(* Logix 5000 project; controller TFF vendor 1 type 14 code 107 rev 34.11; software revision 34.03; part 21 of 36 *)
(* tags used below, declared in another part *)
   Address : DINT;   // Temp Address
   Config : Configuration;   // Index Array used in configuration routines
   AI101 : ALIAS FOR AnalogPoint[10];   // Filtrate Conductivity
   AlarmAnalog : AlarmAnalog[50];   // Analog Alarm Array
   AnalogOutput : AnalogOutput[25];   // Analog Output Array
   AnalogPoint : AnalogInput[50];   // Analog Input Array
   Concentration : Concentration;
   ControlLoop : ControlLoop[20];   // Control Loop Array
   ControlLoop_FeedBagLevel : ALIAS FOR ControlLoop[2];   // Feed Bag Level Control Loop
   ControlLoop_FeedPump : ALIAS FOR ControlLoop[1];   // Feed Pump Control Loop
   Diafiltration : Diafiltration;
   DigitalPoint : DigitalPoint[150];   // Digital Point Array
   Drive : Drive[11];   // Drives Array
   FI003 : ALIAS FOR AnalogPoint[17];
   FlowPath : FlowPath[64];   // Flow Path Array
   FlowPathControl : FlowPathControl;   // Flow Path Control
   FQ_Conc : ALIAS FOR Totalizer[0];   // Concentration Totalizer
   FQ_Diaf : ALIAS FOR Totalizer[1];   // DiafiltrationTotalizer
   Mixer : Mixer;   // Mixer config. structure
   Options : Options;   // Options List
   PCV001 : ALIAS FOR AnalogPoint[3];   // Retentate Pressure Control Valve Position
   PCV101 : ALIAS FOR AnalogPoint[4];   // Filtrate Pressure Control Valve Position
   Phase : Phases[6];   // Phase Control Array
   Phase0_Totalizer_Feed : ALIAS FOR PhaseTotalizer[0];   // Phase 0 Total Feed
   Phase0_Totalizer_Filtrate : ALIAS FOR PhaseTotalizer[6];   // Phase 0 Total Filtrate
   Phase0_Totalizer_Retentate : ALIAS FOR PhaseTotalizer[12];   // Phase 0 Total Retentate
   Phase1_Totalizer_Feed : ALIAS FOR PhaseTotalizer[1];   // Phase 1 Total Feed
   Phase1_Totalizer_Filtrate : ALIAS FOR PhaseTotalizer[7];   // Phase 1 Total Filtrate
   Phase1_Totalizer_Retentate : ALIAS FOR PhaseTotalizer[13];   // Phase 1 Total Retentate
   Phase2_Totalizer_Feed : ALIAS FOR PhaseTotalizer[2];   // Phase 2 Total Feed
   Phase2_Totalizer_Filtrate : ALIAS FOR PhaseTotalizer[8];   // Phase 2 Total Filtrate
   Phase2_Totalizer_Retentate : ALIAS FOR PhaseTotalizer[14];   // Phase 2 Total Retentate
   Phase3_Totalizer_Feed : ALIAS FOR PhaseTotalizer[3];   // Phase 3 Total Feed
   Phase3_Totalizer_Filtrate : ALIAS FOR PhaseTotalizer[9];   // Phase 3 Total Filtrate
   Phase3_Totalizer_Retentate : ALIAS FOR PhaseTotalizer[15];   // Phase 3 Total Retentate
   Phase4_Totalizer_Feed : ALIAS FOR PhaseTotalizer[4];   // Phase 4 Total Feed
   Phase4_Totalizer_Filtrate : ALIAS FOR PhaseTotalizer[10];   // Phase 4 Total Filtrate
   Phase4_Totalizer_Retentate : ALIAS FOR PhaseTotalizer[16];   // Phase 4 Total Retentate
   Phase5_Totalizer_Feed : ALIAS FOR PhaseTotalizer[5];   // Phase 5 Total Feed
   Phase5_Totalizer_Filtrate : ALIAS FOR PhaseTotalizer[11];   // Phase 5 Total Filtrate
   Phase5_Totalizer_Retentate : ALIAS FOR PhaseTotalizer[17];   // Phase 5 Total Retentate
   Rack_Murr_Node4_Instrum_TFF1 : IO_Station;   // Status of Node 4 Instrum TFF1
   Rack_Murr_Node4_Instrum_TFF2 : IO_Station;   // Status of Node 4 Instrum TFF2
   Rack_Murr_Node4_Instrum_TFF3 : IO_Station;   // Status of Node 4 Instrum TFF3
   Rack_Murr_Node4_Instrum_TFF4 : IO_Station;   // Status of Node 4 Instrum TFF4
   Rack_Murr_Node4_Instrum_TFF5 : IO_Station;   // Status of Node 4 Instrum TFF5
   Rack_Murr_Node5_Tank100 : IO_Station;   // Status of Node 5 Tank 100L
   Rack_Murr_Node5_Tank250 : IO_Station;   // Status of Node 5 Tank 250L
   Rack_Murr_Node5_Tank50 : IO_Station;   // Status of Node 5 Tank 50L
   SIC001 : ALIAS FOR Drive[1];   // Feed Pump
   SIC002 : ALIAS FOR Drive[2];   // Transfer Pump
   SIC003 : ALIAS FOR Drive[3];   // Mixer
   SysControl : SysControl;   // General system status and command
   Tank : TankManagement;   // Tank Management
   ThisSystem : SystemType;
   Valve : Valve[100];   // Valve Array
   ValveControl : ValveControl;   // Valve Control
   XV001 : ALIAS FOR Valve[0];   // XV001
   XV002 : ALIAS FOR Valve[1];   // XV002
   XV003 : ALIAS FOR Valve[2];   // XV003
   XV004 : ALIAS FOR Valve[3];   // XV004
   XV005 : ALIAS FOR Valve[4];   // XV005
   XV006 : ALIAS FOR Valve[19];
   XV007 : ALIAS FOR Valve[20];
   XV102 : ALIAS FOR Valve[5];   // XV102
   XV401 : ALIAS FOR Valve[6];   // XV401
   XV402 : ALIAS FOR Valve[7];   // XV402
   XV403 : ALIAS FOR Valve[15];
   XV404 : ALIAS FOR Valve[16];
   XV405 : ALIAS FOR Valve[17];
   XV406 : ALIAS FOR Valve[18];
   XV411 : ALIAS FOR Valve[8];   // XV411
   XV421 : ALIAS FOR Valve[9];   // XV421
   XV431 : ALIAS FOR Valve[10];   // XV431
   XV441 : ALIAS FOR Valve[11];   // XV441
   XV501 : ALIAS FOR Valve[12];   // XV501
   XV502 : ALIAS FOR Valve[13];   // XV502
   XV901 : ALIAS FOR Valve[14];   // XV901
(* Process, continued *)

ROUTINE Config_Drive   (* structured text *)
   (* ==========================================================
   	Config Drive : Configure Drive Structure (for Pumps)
   
   	List of treatments
   		- Drive[1] : Feed Pump SIC001
   		- Drive[2] : Transfer Pump SIC002
   		- Drive[3] : Mixer SIC003
   		- Reset Loop : Set to 0 the Drive[0 and 4 to 10].EnableCfg
   
   -----------------------------------------------------------------------------------------------------------------------------------------------------
   	History
   		2019-AUG-13 - ACTEMIUM - B. Roch - Initial version for Candidate Release 3.00.00.00.a
   ============================================================*)
   
   
   (*Drive[1] : Feed Pump SIC001
   ============================================================*)
   Config.IndexDr := 1 ;
   Drive[1].EnableCfg := 1 ;
   Drive[1].OutputAddress := 3 ;
   Drive[1].InputAddress := 0 ;
   Drive[1].RunInput := 0 ;
   Drive[1].InterlockTimer.PRE := 1000 ;
   Drive[1].ReverseCfg := 0 ;
   Drive[1].DirectionAddress := 0 ;
   
   (*Drive[2] : Transfer Pump SIC002
   ============================================================*)
   Drive[2].EnableCfg := 1 ;
   Drive[2].OutputAddress := 4 ;
   Drive[2].InputAddress := 0 ;
   Drive[2].RunInput := 0 ;
   Drive[2].InterlockTimer.PRE := 1000 ;
   Drive[2].ReverseCfg := 0 ;
   Drive[2].DirectionAddress := 0 ;
   
   (*Drive[3] : Mixer SIC003
   ============================================================*)
   Drive[3].EnableCfg := 1 ;
   Drive[3].OutputAddress := 6 ;
   Drive[3].InputAddress := 0 ;
   Drive[3].RunInput := 0 ;
   Drive[3].InterlockTimer.PRE := 1000 ;
   Drive[3].ReverseCfg := 0 ;
   Drive[3].DirectionAddress := 0 ;
   
   (*Reset Loop : Set to 0 the Drive[0 and 4 to 10].EnableCfg
   ============================================================*)
   for Config.IndexDr := 0 to 10 by 1 do
   	if Config.IndexDr = 0 or Config.IndexDr >= 4 then
   		Drive[Config.IndexDr].EnableCfg := 0 ;
   	End_if ;
   End_for ;
END_ROUTINE

ROUTINE Config_Flowpath   (* structured text *)
   (* =======================================================================
   	Config Flowpath : Configure predifined flowpath
   
   	List of treatments
   		- Critical
   		- Inlets
   		- Flush
   		- Drain
   		- Process
   		- Product Recovery
   		- Open All Main Valve
   		- Close All Main Valve
   		- Open All Valve (reserved)
   		- Close All Valve (reserved)
   		- Reset Loop : Set to 0 the mask and truth of Flowpath[36 to 60]
   
   -----------------------------------------------------------------------------------------------------------------------------------------------------
   	History
   		2019-AUG-13 - ACTEMIUM - B. Roch - Initial version for Candidate Release 3.00.00.00.a
   		2019-SEP-09 - ACTEMIUM - Q. Spindler - Modifications for Candidate Release 3.00.00.00.c
   					- Remove Flush and Drain from the Open all valve and close all valves Flowpath
   		2020-SEP-30 - Merck - Q.Spindler - Modifications for Candidate Release 3.00.00.01.a
   					- Modify flowpath for Closed flowpath option
   					- Add Flexware installation flowpath
   		2023-MAR-03 - Merck - Q.Spindler - Modifications for Candidate Release 3.02.00.00.a
   					- Add Remove TF3S/Closed FP Valves from masks if not enabled
   =========================================================================*)
   
   (* Max flowpath number use as terminal value in loop
   =========================================================================*)
   FlowPathControl.MaxFlowPath := 63 ;
   
   (* Critical
   =========================================================================*)
   (* Critical *)
   
   	FlowPath[2].Mask1 := 2097151 ;
   	FlowPath[2].Mask2 := 0 ;
   	FlowPath[2].Mask3 := 0 ;
   	FlowPath[2].Mask4 := 0 ;
   	FlowPath[2].DrainMask := 1 ;
   	FlowPath[2].FlushMask := 1 ;
   	FlowPath[2].Truth1 := 524299 ;
   	FlowPath[2].Truth2 := 0 ;
   	FlowPath[2].Truth3 := 0 ;
   	FlowPath[2].Truth4 := 0 ;
   	FlowPath[2].DrainTruth := 0 ;
   	FlowPath[2].FlushTruth := 0 ;
   
   
   (* Inlets
   =========================================================================*)
   	(* All Source Valves Open *)
   	FlowPath[3].Mask1 := 1052608 ;
   	FlowPath[3].Mask2 := 0 ;
   	FlowPath[3].Mask3 := 0 ;
   	FlowPath[3].Mask4 := 0 ;
   	FlowPath[3].DrainMask := 0 ;
   	FlowPath[3].FlushMask := 0 ;
   	FlowPath[3].Truth1 := 1052608 ;
   	FlowPath[3].Truth2 := 0 ;
   	FlowPath[3].Truth3 := 0 ;
   	FlowPath[3].Truth4 := 0 ;
   	FlowPath[3].DrainTruth := 0 ;
   	FlowPath[3].FlushTruth := 0 ;
   
   	(* All Source Valves Closed *)
   	FlowPath[4].Mask1 := 1052608 ;
   	FlowPath[4].Mask2 := 0 ;
   	FlowPath[4].Mask3 := 0 ;
   	FlowPath[4].Mask4 := 0 ;
   	FlowPath[4].DrainMask := 0 ;
   	FlowPath[4].FlushMask := 0 ;
   	FlowPath[4].Truth1 := 0 ;
   	FlowPath[4].Truth2 := 0 ;
   	FlowPath[4].Truth3 := 0 ;
   	FlowPath[4].Truth4 := 0 ;
   	FlowPath[4].DrainTruth := 0 ;
   	FlowPath[4].FlushTruth := 0 ;
   
   	(* Feed Source Open *)
   	FlowPath[5].Mask1 := 2068416 ;
   	FlowPath[5].Mask2 := 0 ;
   	FlowPath[5].Mask3 := 0 ;
   	FlowPath[5].Mask4 := 0 ;
   	FlowPath[5].DrainMask := 0 ;
   	FlowPath[5].FlushMask := 0 ;
   	FlowPath[5].Truth1 := 256 ;
   	FlowPath[5].Truth2 := 0 ;
   	FlowPath[5].Truth3 := 0 ;
   	FlowPath[5].Truth4 := 0 ;
   	FlowPath[5].DrainTruth := 0 ;
   	FlowPath[5].FlushTruth := 0 ;
   
   	(* Buffer Source Open *)
   	FlowPath[6].Mask1 := 2068416 ;
   	FlowPath[6].Mask2 := 0 ;
   	FlowPath[6].Mask3 := 0 ;
   	FlowPath[6].Mask4 := 0 ;
   	FlowPath[6].DrainMask := 0 ;
   	FlowPath[6].FlushMask := 0 ;
   	FlowPath[6].Truth1 := 576 ;
   	FlowPath[6].Truth2 := 0 ;
   	FlowPath[6].Truth3 := 0 ;
   	FlowPath[6].Truth4 := 0 ;
   	FlowPath[6].DrainTruth := 0 ;
   	FlowPath[6].FlushTruth := 0 ;
   
   	(* Caustic Source Open *)
   	FlowPath[7].Mask1 := 2068416 ;
   	FlowPath[7].Mask2 := 0 ;
   	FlowPath[7].Mask3 := 0 ;
   	FlowPath[7].Mask4 := 0 ;
   	FlowPath[7].DrainMask := 0 ;
   	FlowPath[7].FlushMask := 0 ;
   	FlowPath[7].Truth1 := 1088 ;
   	FlowPath[7].Truth2 := 0 ;
   	FlowPath[7].Truth3 := 0 ;
   	FlowPath[7].Truth4 := 0 ;
   	FlowPath[7].DrainTruth := 0 ;
   	FlowPath[7].FlushTruth := 0 ;
   
   	(* Water Source Open *)
   	FlowPath[8].Mask1 := 2068416 ;
   	FlowPath[8].Mask2 := 0 ;
   	FlowPath[8].Mask3 := 0 ;
   	FlowPath[8].Mask4 := 0 ;
   	FlowPath[8].DrainMask := 0 ;
   	FlowPath[8].FlushMask := 0 ;
   	FlowPath[8].Truth1 := 2112 ;
   	FlowPath[8].Truth2 := 0 ;
   	FlowPath[8].Truth3 := 0 ;
   	FlowPath[8].Truth4 := 0 ;
   	FlowPath[8].DrainTruth := 0 ;
   	FlowPath[8].FlushTruth := 0 ;
   
   	(* Air Source Open *)
   	FlowPath[9].Mask1 := 2068416 ;
   	FlowPath[9].Mask2 := 0 ;
   	FlowPath[9].Mask3 := 0 ;
   	FlowPath[9].Mask4 := 0 ;
   	FlowPath[9].DrainMask := 0 ;
   	FlowPath[9].FlushMask := 0 ;
   	FlowPath[9].Truth1 := 192 ;
   	FlowPath[9].Truth2 := 0 ;
   	FlowPath[9].Truth3 := 0 ;
   	FlowPath[9].Truth4 := 0 ;
   	FlowPath[9].DrainTruth := 0 ;
   	FlowPath[9].FlushTruth := 0 ;
   
   
   	(* Flush
   =========================================================================*)
   	(* Single Pass Flush (from inlet manifold) *)
   	FlowPath[10].Mask1 := 1044543 ;
   	FlowPath[10].Mask2 := 0 ;
   	FlowPath[10].Mask3 := 0 ;
   	FlowPath[10].Mask4 := 0 ;
   	FlowPath[10].DrainMask := 1 ;
   	FlowPath[10].FlushMask := 1 ;
   	FlowPath[10].Truth1 := 393227 ;
   	FlowPath[10].Truth2 := 0 ;
   	FlowPath[10].Truth3 := 0 ;
   	FlowPath[10].Truth4 := 0 ;
   	FlowPath[10].DrainTruth := 1 ;
   	FlowPath[10].FlushTruth := 1 ;
   
   	(* Single Pass Flush (from recycle bag) *)
   	FlowPath[11].Mask1 := 1044543 ;
   	FlowPath[11].Mask2 := 0 ;
   	FlowPath[11].Mask3 := 0 ;
   	FlowPath[11].Mask4 := 0 ;
   	FlowPath[11].DrainMask := 1 ;
   	FlowPath[11].FlushMask := 1 ;
   	FlowPath[11].Truth1 := 65547 ;
   	FlowPath[11].Truth2 := 0 ;
   	FlowPath[11].Truth3 := 0 ;
   	FlowPath[11].Truth4 := 0 ;
   	FlowPath[11].DrainTruth := 1 ;
   	FlowPath[11].FlushTruth := 0 ;
   
   
   	(* Drain
   =========================================================================*)
   	(* System Drain (without recycle bag) *)
   	FlowPath[12].Mask1 := 1044543 ;
   	FlowPath[12].Mask2 := 0 ;
   	FlowPath[12].Mask3 := 0 ;
   	FlowPath[12].Mask4 := 0 ;
   	FlowPath[12].DrainMask := 1 ;
   	FlowPath[12].FlushMask := 1 ;
   	FlowPath[12].Truth1 := 409647 ;
   	FlowPath[12].Truth2 := 0 ;
   	FlowPath[12].Truth3 := 0 ;
   	FlowPath[12].Truth4 := 0 ;
   	FlowPath[12].DrainTruth := 1 ;
   	FlowPath[12].FlushTruth := 1 ;
   
   	(* System Drain (from recycle bag) *)
   	FlowPath[13].Mask1 := 1044543 ;
   	FlowPath[13].Mask2 := 0 ;
   	FlowPath[13].Mask3 := 0 ;
   	FlowPath[13].Mask4 := 0 ;
   	FlowPath[13].DrainMask := 1 ;
   	FlowPath[13].FlushMask := 1 ;
   	FlowPath[13].Truth1 := 81983 ;
   	FlowPath[13].Truth2 := 0 ;
   	FlowPath[13].Truth3 := 0 ;
   	FlowPath[13].Truth4 := 0 ;
   	FlowPath[13].DrainTruth := 1 ;
   	FlowPath[13].FlushTruth := 0 ;
   
   
   	(* Process
   =========================================================================*)
   	(* Membrane Soak *)
   	FlowPath[14].Mask1 := 1044543 ;
   	FlowPath[14].Mask2 := 0 ;
   	FlowPath[14].Mask3 := 0 ;
   	FlowPath[14].Mask4 := 0 ;
   	FlowPath[14].DrainMask := 1 ;
   	FlowPath[14].FlushMask := 1 ;
   	FlowPath[14].Truth1 := 65539 ;
   	FlowPath[14].Truth2 := 0 ;
   	FlowPath[14].Truth3 := 0 ;
   	FlowPath[14].Truth4 := 0 ;
   	FlowPath[14].DrainTruth := 0 ;
   	FlowPath[14].FlushTruth := 0 ;
   
   	(* Integrity Test *)
   	FlowPath[15].Mask1 := 1044543 ;
   	FlowPath[15].Mask2 := 0 ;
   	FlowPath[15].Mask3 := 0 ;
   	FlowPath[15].Mask4 := 0 ;
   	FlowPath[15].DrainMask := 1 ;
   	FlowPath[15].FlushMask := 1 ;
   	FlowPath[15].Truth1 := 48 ;
   	FlowPath[15].Truth2 := 0 ;
   	FlowPath[15].Truth3 := 0 ;
   	FlowPath[15].Truth4 := 0 ;
   	FlowPath[15].DrainTruth := 0 ;
   	FlowPath[15].FlushTruth := 0 ;
   
   	(* Recycle Bag Fill *)
   	FlowPath[16].Mask1 := 1044543 ;
   	FlowPath[16].Mask2 := 0 ;
   	FlowPath[16].Mask3 := 0 ;
   	FlowPath[16].Mask4 := 0 ;
   	FlowPath[16].DrainMask := 1 ;
   	FlowPath[16].FlushMask := 1 ;
   	FlowPath[16].Truth1 := 524312 ;
   	FlowPath[16].Truth2 := 0 ;
   	FlowPath[16].Truth3 := 0 ;
   	FlowPath[16].Truth4 := 0 ;
   	FlowPath[16].DrainTruth := 0 ;
   	FlowPath[16].FlushTruth := 0 ;
   
   	(* Recycle Bag Drain *)
   	FlowPath[17].Mask1 := 1044543 ;
   	FlowPath[17].Mask2 := 0 ;
   	FlowPath[17].Mask3 := 0 ;
   	FlowPath[17].Mask4 := 0 ;
   	FlowPath[17].DrainMask := 1 ;
   	FlowPath[17].FlushMask := 1 ;
   	FlowPath[17].Truth1 := 81925 ;
   	FlowPath[17].Truth2 := 0 ;
   	FlowPath[17].Truth3 := 0 ;
   	FlowPath[17].Truth4 := 0 ;
   	FlowPath[17].DrainTruth := 0 ;
   	FlowPath[17].FlushTruth := 0 ;
   
   	(* Recovery Filter Flush *)
   	FlowPath[18].Mask1 := 1044543 ;
   	FlowPath[18].Mask2 := 0 ;
   	FlowPath[18].Mask3 := 0 ;
   	FlowPath[18].Mask4 := 0 ;
   	FlowPath[18].DrainMask := 1 ;
   	FlowPath[18].FlushMask := 1 ;
   	FlowPath[18].Truth1 := 65541 ;
   	FlowPath[18].Truth2 := 0 ;
   	FlowPath[18].Truth3 := 0 ;
   	FlowPath[18].Truth4 := 0 ;
   	FlowPath[18].DrainTruth := 0 ;
   	FlowPath[18].FlushTruth := 0 ;
   
   	(* Batch UF or Membrane Recycle *)
   	FlowPath[19].Mask1 := 1044543 ;
   	FlowPath[19].Mask2 := 0 ;
   	FlowPath[19].Mask3 := 0 ;
   	FlowPath[19].Mask4 := 0 ;
   	FlowPath[19].DrainMask := 1 ;
   	FlowPath[19].FlushMask := 1 ;
   	FlowPath[19].Truth1 := 589835 ;
   	FlowPath[19].Truth2 := 0 ;
   	FlowPath[19].Truth3 := 0 ;
   	FlowPath[19].Truth4 := 0 ;
   	FlowPath[19].DrainTruth := 0 ;
   	FlowPath[19].FlushTruth := 0 ;
   
   	(* Fed Batch UF or Diafiltration *)
   	FlowPath[20].Mask1 := 1044543 ;
   	FlowPath[20].Mask2 := 0 ;
   	FlowPath[20].Mask3 := 0 ;
   	FlowPath[20].Mask4 := 0 ;
   	FlowPath[20].DrainMask := 1 ;
   	FlowPath[20].FlushMask := 1 ;
   	FlowPath[20].Truth1 := 589851 ;
   	FlowPath[20].Truth2 := 0 ;
   	FlowPath[20].Truth3 := 0 ;
   	FlowPath[20].Truth4 := 0 ;
   	FlowPath[20].DrainTruth := 0 ;
   	FlowPath[20].FlushTruth := 0 ;
   
   
   	(* Product Recovery
   =========================================================================*)
   	(* Product Recovery 1&3 - Empty Recycle Bag (TF2S) *)
   	FlowPath[21].Mask1 := 1032255 ;
   	FlowPath[21].Mask2 := 0 ;
   	FlowPath[21].Mask3 := 0 ;
   	FlowPath[21].Mask4 := 0 ;
   	FlowPath[21].DrainMask := 1 ;
   	FlowPath[21].FlushMask := 1 ;
   	FlowPath[21].Truth1 := 65541 ;
   	FlowPath[21].Truth2 := 0 ;
   	FlowPath[21].Truth3 := 0 ;
   	FlowPath[21].Truth4 := 0 ;
   	FlowPath[21].DrainTruth := 0 ;
   	FlowPath[21].FlushTruth := 0 ;
   
   	(* Product Recovery 2 - Empty Retentate Line (TF2S) *)
   	FlowPath[22].Mask1 := 1032255 ;
   	FlowPath[22].Mask2 := 0 ;
   	FlowPath[22].Mask3 := 0 ;
   	FlowPath[22].Mask4 := 0 ;
   	FlowPath[22].DrainMask := 1 ;
   	FlowPath[22].FlushMask := 1 ;
   	FlowPath[22].Truth1 := 524312 ;
   	FlowPath[22].Truth2 := 0 ;
   	FlowPath[22].Truth3 := 0 ;
   	FlowPath[22].Truth4 := 0 ;
   	FlowPath[22].DrainTruth := 0 ;
   	FlowPath[22].FlushTruth := 0 ;
   
   	(* Product Recovery 4 - Empty Membranes (TF2S) *)
   	FlowPath[23].Mask1 := 1032255 ;
   	FlowPath[23].Mask2 := 0 ;
   	FlowPath[23].Mask3 := 0 ;
   	FlowPath[23].Mask4 := 0 ;
   	FlowPath[23].DrainMask := 1 ;
   	FlowPath[23].FlushMask := 1 ;
   	FlowPath[23].Truth1 := 22 ;
   	FlowPath[23].Truth2 := 0 ;
   	FlowPath[23].Truth3 := 0 ;
   	FlowPath[23].Truth4 := 0 ;
   	FlowPath[23].DrainTruth := 0 ;
   	FlowPath[23].FlushTruth := 0 ;
   
   	(* Product Recovery 1&5 - Empty Recycle Bag (TF3S) *)
   	FlowPath[24].Mask1 := 1044543 ;
   	FlowPath[24].Mask2 := 0 ;
   	FlowPath[24].Mask3 := 0 ;
   	FlowPath[24].Mask4 := 0 ;
   	FlowPath[24].DrainMask := 1 ;
   	FlowPath[24].FlushMask := 1 ;
   	FlowPath[24].Truth1 := 65541 ;
   	FlowPath[24].Truth2 := 0 ;
   	FlowPath[24].Truth3 := 0 ;
   	FlowPath[24].Truth4 := 0 ;
   	FlowPath[24].DrainTruth := 0 ;
   	FlowPath[24].FlushTruth := 0 ;
   
   	(* Product Recovery 2 - Empty Membranes (TF3S) *)
   	FlowPath[25].Mask1 := 1044543 ;
   	FlowPath[25].Mask2 := 0 ;
   	FlowPath[25].Mask3 := 0 ;
   	FlowPath[25].Mask4 := 0 ;
   	FlowPath[25].DrainMask := 1 ;
   	FlowPath[25].FlushMask := 1 ;
   	FlowPath[25].Truth1 := 22 ;
   	FlowPath[25].Truth2 := 0 ;
   	FlowPath[25].Truth3 := 0 ;
   	FlowPath[25].Truth4 := 0 ;
   	FlowPath[25].DrainTruth := 0 ;
   	FlowPath[25].FlushTruth := 0 ;
   
   	(* Product Recovery 3&6 - Empty Bypass (TF3S) *)
   	FlowPath[26].Mask1 := 1044543 ;
   	FlowPath[26].Mask2 := 0 ;
   	FlowPath[26].Mask3 := 0 ;
   	FlowPath[26].Mask4 := 0 ;
   	FlowPath[26].DrainMask := 1 ;
   	FlowPath[26].FlushMask := 1 ;
   	FlowPath[26].Truth1 := 12310 ;
   	FlowPath[26].Truth2 := 0 ;
   	FlowPath[26].Truth3 := 0 ;
   	FlowPath[26].Truth4 := 0 ;
   	FlowPath[26].DrainTruth := 0 ;
   	FlowPath[26].FlushTruth := 0 ;
   
   	(* Product Recovery 4 - Empty Retentate Line (TF3S) *)
   	FlowPath[27].Mask1 := 1044543 ;
   	FlowPath[27].Mask2 := 0 ;
   	FlowPath[27].Mask3 := 0 ;
   	FlowPath[27].Mask4 := 0 ;
   	FlowPath[27].DrainMask := 1 ;
   	FlowPath[27].FlushMask := 1 ;
   	FlowPath[27].Truth1 := 524312 ;
   	FlowPath[27].Truth2 := 0 ;
   	FlowPath[27].Truth3 := 0 ;
   	FlowPath[27].Truth4 := 0 ;
   	FlowPath[27].DrainTruth := 0 ;
   	FlowPath[27].FlushTruth := 0 ;
   
   
   (* Open All Main Valve
   =========================================================================*)
   	(* All Main Flowpath Valves Open *)
   	FlowPath[28].Mask1 := 1044543 ;
   	FlowPath[28].Mask2 := 0 ;
   	FlowPath[28].Mask3 := 0 ;
   	FlowPath[28].Mask4 := 0 ;
   	FlowPath[28].DrainMask := 1 ;
   	FlowPath[28].FlushMask := 1 ;
   	FlowPath[28].Truth1 := 606271 ;
   	FlowPath[28].Truth2 := 0 ;
   	FlowPath[28].Truth3 := 0 ;
   	FlowPath[28].Truth4 := 0 ;
   	FlowPath[28].DrainTruth := 0 ;
   	FlowPath[28].FlushTruth := 0 ;
   
   
   (* Close All Main Valve
   =========================================================================*)
   	(* All Main Flowpath Valves Closed *)
   	FlowPath[29].Mask1 := 1044543 ;
   	FlowPath[29].Mask2 := 0 ;
   	FlowPath[29].Mask3 := 0 ;
   	FlowPath[29].Mask4 := 0 ;
   	FlowPath[29].DrainMask := 1 ;
   	FlowPath[29].FlushMask := 1 ;
   	FlowPath[29].Truth1 := 0 ;
   	FlowPath[29].Truth2 := 0 ;
   	FlowPath[29].Truth3 := 0 ;
   	FlowPath[29].Truth4 := 0 ;
   	FlowPath[29].DrainTruth := 0 ;
   	FlowPath[29].FlushTruth := 0 ;
   
   
   (* Flowpath from 30 to 34 are reserved for User *)
   
   	(* FlexWare Installation *)
   	FlowPath[35].Mask1 := 2068416 ;
   	FlowPath[35].Mask2 := 0 ;
   	FlowPath[35].Mask3 := 0 ;
   	FlowPath[35].Mask4 := 0 ;
   	FlowPath[35].DrainMask := 0 ;
   	FlowPath[35].FlushMask := 0 ;
   	FlowPath[35].Truth1 := 2068416 ;
   	FlowPath[35].Truth2 := 0 ;
   	FlowPath[35].Truth3 := 0 ;
   	FlowPath[35].Truth4 := 0 ;
   	FlowPath[35].DrainTruth := 0 ;
   	FlowPath[35].FlushTruth := 0 ;
   
   
   // Remove TF3S Valves from mask if not enabled
   IF NOT Options.TF3S THEN
   	FOR Config.IndexFlowpath := 2 to 29 by 1 do
   		FlowPath[Config.IndexFlowpath].Mask1.12 := 0 ; //XV501
   		FlowPath[Config.IndexFlowpath].Mask1.13 := 0 ; //XV502
   	End_for ;
   		FlowPath[35].Mask1.12 := 0 ; //XV501
   		FlowPath[35].Mask1.13 := 0 ; //XV502
   END_IF;
   
   // Remove Closed FP Valves from mask if not enabled
   IF NOT Options.ClosedFP THEN
   	FOR Config.IndexFlowpath := 2 to 29 by 1 do
   		FlowPath[Config.IndexFlowpath].Mask1.15 := 0 ; //XV403
   		FlowPath[Config.IndexFlowpath].Mask1.16 := 0 ; //XV404
   		FlowPath[Config.IndexFlowpath].Mask1.17 := 0 ; //XV405
   		FlowPath[Config.IndexFlowpath].Mask1.18 := 0 ; //XV406
   		FlowPath[Config.IndexFlowpath].Mask1.19 := 0 ; //XV006
   		FlowPath[Config.IndexFlowpath].Mask1.20 := 0 ; //XV007
   	End_for ;
   		FlowPath[35].Mask1.15 := 0 ; //XV403
   		FlowPath[35].Mask1.16 := 0 ; //XV404
   		FlowPath[35].Mask1.17 := 0 ; //XV405
   		FlowPath[35].Mask1.18 := 0 ; //XV406
   		FlowPath[35].Mask1.19 := 0 ; //XV006
   		FlowPath[35].Mask1.20 := 0 ; //XV007
   END_IF;
   
   
   (* Open All Valve (reserved)
   =========================================================================*)
   (* Open All Valve *)
   FlowPath[61].Mask1 := -1 ;
   FlowPath[61].Mask2 := 0 ;
   FlowPath[61].Mask3 := 0 ;
   FlowPath[61].Mask4 := 0 ;
   FlowPath[61].DrainMask := 0 ;
   FlowPath[61].FlushMask := 0 ;
   FlowPath[61].Truth1 := -1 ;
   FlowPath[61].Truth2 := 0 ;
   FlowPath[61].Truth3 := 0 ;
   FlowPath[61].Truth4 := 0 ;
   FlowPath[61].DrainTruth := 0 ;
   FlowPath[61].FlushTruth := 0 ;
   
   (* Close All Valve (reserved)
   =========================================================================*)
   (* Close All Valve *)
   FlowPath[62].Mask1 := -1 ;
   FlowPath[62].Mask2 := 0 ;
   FlowPath[62].Mask3 := 0 ;
   FlowPath[62].Mask4 := 0 ;
   FlowPath[62].DrainMask := 0 ;
   FlowPath[62].FlushMask := 0 ;
   FlowPath[62].Truth1 := 0 ;
   FlowPath[62].Truth2 := 0 ;
   FlowPath[62].Truth3 := 0 ;
   FlowPath[62].Truth4 := 0 ;
   FlowPath[62].DrainTruth := 0 ;
   FlowPath[62].FlushTruth := 0 ;
   
   (*Reset Loop : Set to 0 the Flowpath[36 to 60]
   ============================================================*)
   FOR Config.IndexFlowpath := 36 to 60 by 1 do
   	FlowPath[Config.IndexFlowpath].Mask1 := 0 ;
   	FlowPath[Config.IndexFlowpath].Mask2 := 0 ;
   	FlowPath[Config.IndexFlowpath].Mask3 := 0 ;
   	FlowPath[Config.IndexFlowpath].Mask4 := 0 ;
   	FlowPath[Config.IndexFlowpath].DrainMask := 0 ;
   	FlowPath[Config.IndexFlowpath].FlushMask := 0 ;
   	FlowPath[Config.IndexFlowpath].Truth1 := 0 ;
   	FlowPath[Config.IndexFlowpath].Truth2 := 0 ;
   	FlowPath[Config.IndexFlowpath].Truth3 := 0 ;
   	FlowPath[Config.IndexFlowpath].Truth4 := 0 ;
   	FlowPath[Config.IndexFlowpath].Status := 0 ;
   	FlowPath[Config.IndexFlowpath].DrainTruth := 0 ;
   	FlowPath[Config.IndexFlowpath].FlushTruth := 0 ;
   End_for ;
END_ROUTINE

ROUTINE Config_Options   (* structured text *)
   (* ==========================================================
   	Config Options : Configure Options
   
   	List of treatments
   		- Configure Instrum TFF options
   		- Configure Tank options
   		- Configure Flag for current installed clamshell
   
   -----------------------------------------------------------------------------------------------------------------------------------------------------
   	History
   		2019-AUG-13 - ACTEMIUM - B. Roch - Initial version for Candidate Release 3.00.00.00.a
   ============================================================*)
   
   (*Configure options if option Simulation mode is disabled*)
   If Not SysControl.Simulate_Options Then
   
   	(* Configure Instrum TFF options
   	Set options depending on which INSTRUM_TFF I/O device is active
   	============================================================*)
   
   	(*No Device Connected*)
   	IF NOT Rack_Murr_Node4_Instrum_TFF1.Node_Comm_Status AND NOT Rack_Murr_Node4_Instrum_TFF2.Node_Comm_Status AND NOT Rack_Murr_Node4_Instrum_TFF3.Node_Comm_Status AND NOT Rack_Murr_Node4_Instrum_TFF4.Node_Comm_Status AND NOT Rack_Murr_Node4_Instrum_TFF5.Node_Comm_Status THEN
   	Options.No_Device_Connected := 1 ;
   	Options.AI102_AI103 := 0 ;
   	Options.AI101 := 0 ;
   	Options.AI101_AI102_AI103 := 0 ;
   	Options.AI101_AI104 := 0 ;
   	Options.AI101_AI102_AI103_AI104 := 0 ;
   	END_IF;
   
   	(*UV Probe Device*)
   	IF Rack_Murr_Node4_Instrum_TFF1.Node_Comm_Status THEN
   	Options.No_Device_Connected := 0 ;
   	Options.AI102_AI103 := 1 ;
   	Options.AI101 := 0 ;
   	Options.AI101_AI102_AI103 := 0 ;
   	Options.AI101_AI104 := 0 ;
   	Options.AI101_AI102_AI103_AI104 := 0 ;
   	END_IF;
   
   	(*Conductivity*)
   	IF Rack_Murr_Node4_Instrum_TFF2.Node_Comm_Status THEN
   	Options.No_Device_Connected := 0 ;
   	Options.AI102_AI103 := 0 ;
   	Options.AI101 := 1 ;
   	Options.AI101_AI102_AI103 := 0 ;
   	Options.AI101_AI104 := 0 ;
   	Options.AI101_AI102_AI103_AI104 := 0 ;
   	END_IF;
   
   	(*UV and Conductivity*)
   	IF Rack_Murr_Node4_Instrum_TFF3.Node_Comm_Status THEN
   	Options.No_Device_Connected := 0 ;
   	Options.AI102_AI103 := 0 ;
   	Options.AI101 := 0 ;
   	Options.AI101_AI102_AI103 := 1 ;
   	Options.AI101_AI104 := 0 ;
   	Options.AI101_AI102_AI103_AI104 := 0 ;
   	END_IF;
   
   	(*Conductivity and pH*)
   	IF Rack_Murr_Node4_Instrum_TFF4.Node_Comm_Status THEN
   	Options.No_Device_Connected := 0 ;
   	Options.AI102_AI103 := 0 ;
   	Options.AI101 := 0 ;
   	Options.AI101_AI102_AI103 := 0 ;
   	Options.AI101_AI104 := 1 ;
   	Options.AI101_AI102_AI103_AI104 := 0 ;
   	END_IF;
   
   	(*UV and Conductivity and pH*)
   	IF Rack_Murr_Node4_Instrum_TFF5.Node_Comm_Status THEN
   	Options.No_Device_Connected := 0 ;
   	Options.AI102_AI103 := 0 ;
   	Options.AI101 := 0 ;
   	Options.AI101_AI102_AI103 := 0 ;
   	Options.AI101_AI104 := 0 ;
   	Options.AI101_AI102_AI103_AI104 := 1 ;
   	END_IF;
   
   	(* Configure Tank options
   	Set options depending on which TANK I/O device is active
   	============================================================*)
   
   	(*No Tank Connected*)
   	IF NOT Rack_Murr_Node5_Tank50.Node_Comm_Status AND NOT Rack_Murr_Node5_Tank100.Node_Comm_Status AND NOT Rack_Murr_Node5_Tank250.Node_Comm_Status THEN
   	Options.No_Tank := 1 ;
   	Options.Tank50 := 0 ;
   	Options.Tank100 := 0 ;
   	Options.Tank250 := 0 ;
   	Tank.Config.Option_Current := 0 ;
   	END_IF;
   
   	(*Tank 50*)
   	IF Rack_Murr_Node5_Tank50.Node_Comm_Status THEN
   	Options.No_Tank := 0 ;
   	Options.Tank50 := 1 ;
   	Options.Tank100 := 0 ;
   	Options.Tank250 := 0 ;
   	Tank.Config.Option_Current := 1 ;
   	END_IF;
   
   	(*Tank 100*)
   	IF Rack_Murr_Node5_Tank100.Node_Comm_Status THEN
   	Options.No_Tank := 0 ;
   	Options.Tank50 := 0 ;
   	Options.Tank100 := 1 ;
   	Options.Tank250 := 0 ;
   	Tank.Config.Option_Current := 2 ;
   	END_IF;
   
   	(*Tank 250*)
   	IF Rack_Murr_Node5_Tank250.Node_Comm_Status THEN
   	Options.No_Tank := 0 ;
   	Options.Tank50 := 0 ;
   	Options.Tank100 := 0 ;
   	Options.Tank250 := 1 ;
   	Tank.Config.Option_Current := 3 ;
   	END_IF;
   
   End_If;
   
   
   (*Simulate Tank Range*)
   IF Tank.Config.Simulate THEN
   
   	CASE	Tank.Config.Option_Simulate OF
   		0:	Options.No_Tank := 1 ;
   			Options.Tank50 := 0 ;
   			Options.Tank100 := 0 ;
   			Options.Tank250 := 0 ;
   			Tank.Config.Option_Current := 0 ;
   		1:	Options.No_Tank := 0 ;
   			Options.Tank50 := 1 ;
   			Options.Tank100 := 0 ;
   			Options.Tank250 := 0 ;
   			Tank.Config.Option_Current := 1 ;
   		2:	Options.No_Tank := 0 ;
   			Options.Tank50 := 0 ;
   			Options.Tank100 := 1 ;
   			Options.Tank250 := 0 ;
   			Tank.Config.Option_Current := 2 ;
   		3:	Options.No_Tank := 0 ;
   			Options.Tank50 := 0 ;
   			Options.Tank100 := 0 ;
   			Options.Tank250 := 1 ;
   			Tank.Config.Option_Current := 3 ;
   	ELSE 	Options.No_Tank := 1 ;
   			Options.Tank50 := 0 ;
   			Options.Tank100 := 0 ;
   			Options.Tank250 := 0 ;
   			Tank.Config.Option_Current := 0 ;
   	END_CASE;
   
   END_IF;
   
   (* Configure Flag for current installed clamshell
   Used to create the CCP Configuration file based on current clamshell
   ============================================================*)
   IF ThisSystem.MoldType = 123 THEN
   
   	Options.TF2S := 1 ;
   	Options.TF3S := 0 ;
   
   ELSIF ThisSystem.MoldType = 124 THEN
   
   	Options.TF3S := 1 ;
   	Options.TF2S := 0 ;
   
   END_IF;
END_ROUTINE

ROUTINE Config_Reset   (* structured text *)
// Set to 0  all settings
   (* ==========================================================
   	Config Reset : 	When config.reset command is activated,AnalogPoint, AlarmAnalog, AnalogOutput, Drive, DigitalPoint and Valve structure
   					are initialized to 0.
   
   	List of treatments
   		- AnalogPoint Structure reset [0] to [49]
   		- AlarmAnalog Structure reset [0] to [49]
   		- AnalogOutput Structure reset [0] to [24]
   		- Drive Structure reset [0] to [10]
   		- DigitalPoint Structure reset [0] to [149]
   		- Valve Structure reset [0] to [99]
   
   -----------------------------------------------------------------------------------------------------------------------------------------------------
   	History
   		2019-AUG-13 - ACTEMIUM - B. Roch - Initial version for Candidate Release 3.00.00.00.a
   ============================================================*)
   
   
   (*Structure Reset [0] to [149]
   ============================================================*)
   IF Config.Reset THEN
   	FOR Config.IndexReset := 0 TO 149 BY 1 Do
   		IF Config.IndexReset <= 49 THEN
   		(*AnalogPoint Structure Reset [0] to [49]
   		====================================================*)
   			AnalogPoint[Config.IndexReset].OutofRange := 0 ;
   			AnalogPoint[Config.IndexReset].FilterType := 0 ;
   			AnalogPoint[Config.IndexReset].AveragingTotal := 0 ;
   			AnalogPoint[Config.IndexReset].Address := 0 ;
   			AnalogPoint[Config.IndexReset].RawMin := 0 ;
   			AnalogPoint[Config.IndexReset].RawMax := 0 ;
   			AnalogPoint[Config.IndexReset].RawValue := 0 ;
   			AnalogPoint[Config.IndexReset].RawLowLimit := 0 ;
   			AnalogPoint[Config.IndexReset].RawHighLimit := 0 ;
   			AnalogPoint[Config.IndexReset].FilterUser := 0 ;
   			AnalogPoint[Config.IndexReset].FilteredRaw := 0 ;
   			AnalogPoint[Config.IndexReset].FilterActual := 0 ;
   			AnalogPoint[Config.IndexReset].ScaledMin := 0 ;
   			AnalogPoint[Config.IndexReset].ScaledMax := 0 ;
   			AnalogPoint[Config.IndexReset].RangeMin := 0 ;
   			AnalogPoint[Config.IndexReset].RangeMax := 0 ;
   			AnalogPoint[Config.IndexReset].RangeMinSave := 0 ;
   			AnalogPoint[Config.IndexReset].RangeMaxSave := 0 ;
   			AnalogPoint[Config.IndexReset].RealCfg := 0 ;
   			AnalogPoint[Config.IndexReset].EnableCfg := 0 ;
   			AnalogPoint[Config.IndexReset].OverrideCfg := 0 ;
   
   		(*AlarmAnalog Structure Reset [0] to [49]
   		====================================================*)
   			AlarmAnalog[Config.IndexReset].Override := 0 ;
   			AlarmAnalog[Config.IndexReset].Disable := 0 ;
   			AlarmAnalog[Config.IndexReset].LOLODisable := 0 ;
   			AlarmAnalog[Config.IndexReset].LODisable := 0 ;
   			AlarmAnalog[Config.IndexReset].HIDisable := 0 ;
   			AlarmAnalog[Config.IndexReset].HIHIDisable := 0 ;
   			AlarmAnalog[Config.IndexReset].HIHIEnable := 0 ;
   			AlarmAnalog[Config.IndexReset].FeedPumpEnable := 0 ;
   			AlarmAnalog[Config.IndexReset].FeedPumpTag := 0 ;
   			AlarmAnalog[Config.IndexReset].TransferPumpEnable := 0 ;
   			AlarmAnalog[Config.IndexReset].TransferPumpTag := 0 ;
   			AlarmAnalog[Config.IndexReset].LOLO := 0 ;
   			AlarmAnalog[Config.IndexReset].LO := 0 ;
   			AlarmAnalog[Config.IndexReset].HI := 0 ;
   			AlarmAnalog[Config.IndexReset].HIHI := 0 ;
   			AlarmAnalog[Config.IndexReset].LOLOTimer.PRE := 0 ;
   			AlarmAnalog[Config.IndexReset].LOTimer.PRE := 0 ;
   			AlarmAnalog[Config.IndexReset].HITimer.PRE := 0 ;
   			AlarmAnalog[Config.IndexReset].HIHITimer.PRE := 0 ;
   			AlarmAnalog[Config.IndexReset].EnableCfg := 0 ;
   		End_IF;
   
   		(*AnalogOutput Structure Reset [0] to [24]
   		====================================================*)
   		IF Config.IndexReset <= 24 THEN
   			AnalogOutput[Config.IndexReset].RawValue := 0 ;
   			AnalogOutput[Config.IndexReset].RawMin := 0 ;
   			AnalogOutput[Config.IndexReset].RawMax := 0 ;
   			AnalogOutput[Config.IndexReset].ScaledMin := 0 ;
   			AnalogOutput[Config.IndexReset].ScaledMax := 0 ;
   			AnalogOutput[Config.IndexReset].EnableCfg := 0 ;
   		End_IF;
   
   		(*Drive Structure Reset [0] to [10]
   		====================================================*)
   		IF Config.IndexReset <= 10 THEN
   			Drive[Config.IndexReset].OutputAddress := 0 ;
   			Drive[Config.IndexReset].InputAddress := 0 ;
   			Drive[Config.IndexReset].RunInput := 0 ;
   			Drive[Config.IndexReset].InterlockTimer.PRE := 0 ;
   			Drive[Config.IndexReset].EnableCfg := 0 ;
   			Drive[Config.IndexReset].ReverseCfg := 0 ;
   			Drive[Config.IndexReset].Direction := 0 ;
   			Drive[Config.IndexReset].DirectionAddress := 0 ;
   		End_IF;
   
   		IF Config.IndexReset <= 99 THEN
   				(*Valves Structure Reset [0] to [99]
   		====================================================*)
   		Valve[Config.IndexReset].ZSOpenEnable := 0 ;
   		Valve[Config.IndexReset].ZSCloseEnable := 0 ;
   		Valve[Config.IndexReset].ZSOverride := 0 ;
   		Valve[Config.IndexReset].FailState := 0 ;
   		Valve[Config.IndexReset].Ports := 0 ;
   		Valve[Config.IndexReset].EnableCfg := 0 ;
   		Valve[Config.IndexReset].StatusWord := 0 ;
   		Valve[Config.IndexReset].ZSOpenAddress := 0 ;
   		Valve[Config.IndexReset].ZSCloseAddress := 0 ;
   		Valve[Config.IndexReset].OutputAddress := 0 ;
   		Valve[Config.IndexReset].AlarmTimer.PRE := 0 ;
   		Valve[Config.IndexReset].AutoCloseTimer.PRE := 0 ;
   		End_IF;
   
   		(*DigitalPoint Structure Reset [0] to [149]
   		====================================================*)
   		DigitalPoint[Config.IndexReset].Override := 0 ;
   		DigitalPoint[Config.IndexReset].DelayTimer.PRE := 0 ;
   		DigitalPoint[Config.IndexReset].Priority := 0 ;
   		DigitalPoint[Config.IndexReset].EnableCfg := 0 ;
   		DigitalPoint[Config.IndexReset].ActiveStateCFg := 0 ;
   		DigitalPoint[Config.IndexReset].RealInputCfg := 0 ;
   		DigitalPoint[Config.IndexReset].InputAddressCfg := 0 ;
   		DigitalPoint[Config.IndexReset].AlarmCfg := 0 ;
   		DigitalPoint[Config.IndexReset].AlarmStateCfg := 0 ;
   		DigitalPoint[Config.IndexReset].OverrideCfg := 0 ;
   		DigitalPoint[Config.IndexReset].PriorityCfg := 0 ;
   		DigitalPoint[Config.IndexReset].Cond1Cfg := 0 ;
   		DigitalPoint[Config.IndexReset].Cond2Cfg := 0 ;
   		DigitalPoint[Config.IndexReset].FlashingInputCfg := 0 ;
   
   	END_FOR;
   End_IF;
   (*Reset config.reset to execute routine one time*)
   Config.Reset := 0;
END_ROUTINE

ROUTINE Config_Totalizers   (* structured text *)
   (* ==========================================================
   	Config Totalizers : Configure Totalizers Structure
   
   	List of treatments
   		- Phase 0 Totalizers
   		- Phase 1 Totalizers
   		- Phase 2 Totalizers
   		- Phase 3 Totalizers
   		- Phase 4 Totalizers
   		- Phase 5 Totalizers
   		- Concentration and Diafiltration Totalizers
   
   -----------------------------------------------------------------------------------------------------------------------------------------------------
   	History
   		2019-AUG-13 - ACTEMIUM - B. Roch - Initial version for Candidate Release 3.00.00.00.a
   		2020-SEP-29 - Merck - Q. Spindler - Modifications for Candidate Release 3.00.00.01.a
   					- Add Retentate totalizers
   		2020-NOV-24 - Merck - Q. Spindler - Modifications for Candidate Release 3.00.00.01.b
   					- Change Retentate Flowmeter option
   ============================================================*)
   
   
   (*Phase 0 Totalizers
   ============================================================*)
   Phase0_Totalizer_Feed.EnableCfg := 1 ;
   Phase0_Totalizer_Feed.SourceAddressCfg := 42 ;
   Phase0_Totalizer_Feed.SourceTypeCfg := 0 ;
   Phase0_Totalizer_Feed.PVscale := 60 ;
   
   
   IF Options.No_Filtrate_Measurement THEN
   	Phase0_Totalizer_Filtrate.EnableCfg := 0 ;
   ELSE
   	Phase0_Totalizer_Filtrate.EnableCfg := 1 ;
   END_IF;
   
   Phase0_Totalizer_Filtrate.SourceAddressCfg := 2 ;
   Phase0_Totalizer_Filtrate.SourceTypeCfg := 0 ;
   Phase0_Totalizer_Filtrate.PVscale := 60 ;
   
   IF Options.FI003 THEN
   	Phase0_Totalizer_Retentate.EnableCfg := 1 ;
   ELSE
   	Phase0_Totalizer_Retentate.EnableCfg := 0 ;
   END_IF;
   
   Phase0_Totalizer_Retentate.SourceAddressCfg := 17 ;
   Phase0_Totalizer_Retentate.SourceTypeCfg := 0 ;
   Phase0_Totalizer_Retentate.PVscale := 60 ;
   
   (*Phase 1 Totalizers
   ============================================================*)
   Phase1_Totalizer_Feed.EnableCfg := 1 ;
   Phase1_Totalizer_Feed.SourceAddressCfg := 42 ;
   Phase1_Totalizer_Feed.SourceTypeCfg := 0 ;
   Phase1_Totalizer_Feed.PVscale := 60 ;
   
   IF Options.No_Filtrate_Measurement THEN
   	Phase1_Totalizer_Filtrate.EnableCfg := 0 ;
   ELSE
   	Phase1_Totalizer_Filtrate.EnableCfg := 1 ;
   END_IF;
   
   Phase1_Totalizer_Filtrate.SourceAddressCfg := 2 ;
   Phase1_Totalizer_Filtrate.SourceTypeCfg := 0 ;
   Phase1_Totalizer_Filtrate.PVscale := 60 ;
   
   IF Options.FI003 THEN
   	Phase1_Totalizer_Retentate.EnableCfg := 1 ;
   ELSE
   	Phase1_Totalizer_Retentate.EnableCfg := 0 ;
   END_IF;
   
   Phase1_Totalizer_Retentate.SourceAddressCfg := 17 ;
   Phase1_Totalizer_Retentate.SourceTypeCfg := 0 ;
   Phase1_Totalizer_Retentate.PVscale := 60 ;
   
   (*Phase 2 Totalizers
   ============================================================*)
   Phase2_Totalizer_Feed.EnableCfg := 1 ;
   Phase2_Totalizer_Feed.SourceAddressCfg := 42 ;
   Phase2_Totalizer_Feed.SourceTypeCfg := 0 ;
   Phase2_Totalizer_Feed.PVscale := 60 ;
   
   IF Options.No_Filtrate_Measurement THEN
   	Phase2_Totalizer_Filtrate.EnableCfg := 0 ;
   ELSE
   	Phase2_Totalizer_Filtrate.EnableCfg := 1 ;
   END_IF;
   
   Phase2_Totalizer_Filtrate.SourceAddressCfg := 2 ;
   Phase2_Totalizer_Filtrate.SourceTypeCfg := 0 ;
   Phase2_Totalizer_Filtrate.PVscale := 60 ;
   
   IF Options.FI003 THEN
   	Phase2_Totalizer_Retentate.EnableCfg := 1 ;
   ELSE
   	Phase2_Totalizer_Retentate.EnableCfg := 0 ;
   END_IF;
   
   Phase2_Totalizer_Retentate.SourceAddressCfg := 17 ;
   Phase2_Totalizer_Retentate.SourceTypeCfg := 0 ;
   Phase2_Totalizer_Retentate.PVscale := 60 ;
   
   (*Phase 3 Totalizers
   ============================================================*)
   Phase3_Totalizer_Feed.EnableCfg := 1 ;
   Phase3_Totalizer_Feed.SourceAddressCfg := 42 ;
   Phase3_Totalizer_Feed.SourceTypeCfg := 0 ;
   Phase3_Totalizer_Feed.PVscale := 60 ;
   
   IF Options.No_Filtrate_Measurement THEN
   	Phase3_Totalizer_Filtrate.EnableCfg := 0 ;
   ELSE
   	Phase3_Totalizer_Filtrate.EnableCfg := 1 ;
   END_IF;
   
   Phase3_Totalizer_Filtrate.SourceAddressCfg := 2 ;
   Phase3_Totalizer_Filtrate.SourceTypeCfg := 0 ;
   Phase3_Totalizer_Filtrate.PVscale := 60 ;
   
   IF Options.FI003 THEN
   	Phase3_Totalizer_Retentate.EnableCfg := 1 ;
   ELSE
   	Phase3_Totalizer_Retentate.EnableCfg := 0 ;
   END_IF;
   
   Phase3_Totalizer_Retentate.SourceAddressCfg := 17 ;
   Phase3_Totalizer_Retentate.SourceTypeCfg := 0 ;
   Phase3_Totalizer_Retentate.PVscale := 60 ;
   
   (*Phase 4 Totalizers
   ============================================================*)
   Phase4_Totalizer_Feed.EnableCfg := 1 ;
   Phase4_Totalizer_Feed.SourceAddressCfg := 42 ;
   Phase4_Totalizer_Feed.SourceTypeCfg := 0 ;
   Phase4_Totalizer_Feed.PVscale := 60 ;
   
   IF Options.No_Filtrate_Measurement THEN
   	Phase4_Totalizer_Filtrate.EnableCfg := 0 ;
   ELSE
   	Phase4_Totalizer_Filtrate.EnableCfg := 1 ;
   END_IF;
   
   Phase4_Totalizer_Filtrate.SourceAddressCfg := 2 ;
   Phase4_Totalizer_Filtrate.SourceTypeCfg := 0 ;
   Phase4_Totalizer_Filtrate.PVscale := 60 ;
   
   IF Options.FI003 THEN
   	Phase4_Totalizer_Retentate.EnableCfg := 1 ;
   ELSE
   	Phase4_Totalizer_Retentate.EnableCfg := 0 ;
   END_IF;
   
   Phase4_Totalizer_Retentate.SourceAddressCfg := 17 ;
   Phase4_Totalizer_Retentate.SourceTypeCfg := 0 ;
   Phase4_Totalizer_Retentate.PVscale := 60 ;
   
   (*Phase 5 Totalizers
   ============================================================*)
   Phase5_Totalizer_Feed.EnableCfg := 1 ;
   Phase5_Totalizer_Feed.SourceAddressCfg := 42 ;
   Phase5_Totalizer_Feed.SourceTypeCfg := 0 ;
   Phase5_Totalizer_Feed.PVscale := 60 ;
   
   IF Options.No_Filtrate_Measurement THEN
   	Phase5_Totalizer_Filtrate.EnableCfg := 0 ;
   ELSE
   	Phase5_Totalizer_Filtrate.EnableCfg := 1 ;
   END_IF;
   
   Phase5_Totalizer_Filtrate.SourceAddressCfg := 2 ;
   Phase5_Totalizer_Filtrate.SourceTypeCfg := 0 ;
   Phase5_Totalizer_Filtrate.PVscale := 60 ;
   
   IF Options.FI003 THEN
   	Phase5_Totalizer_Retentate.EnableCfg := 1 ;
   ELSE
   	Phase5_Totalizer_Retentate.EnableCfg := 0 ;
   END_IF;
   
   Phase5_Totalizer_Retentate.SourceAddressCfg := 17 ;
   Phase5_Totalizer_Retentate.SourceTypeCfg := 0 ;
   Phase5_Totalizer_Retentate.PVscale := 60 ;
   
   (*Concentration and Diafiltration Totalizers
   ============================================================*)
   
   FQ_Conc.PVscale := 60 ;
   FQ_Diaf.PVscale := 60 ;
END_ROUTINE

ROUTINE Config_Valve   (* structured text *)
// Apply the default configuration
   (* ==========================================================
   	Config Valve : Configure Valve Structure
   
   	List of treatments
   		- Valve[0] : XV001 Valve XV001
   		- Valve[1] : XV002 Valve XV002
   		- Valve[2] : XV003 Valve XV003
   		- Valve[3] : XV004 Valve XV004
   		- Valve[4] : XV005 Valve XV005
   		- Valve[5] : XV102 Valve XV102
   		- Valve[6] : XV401 Valve XV401
   		- Valve[7] : XV402 Valve XV402
   		- Valve[8] : XV411 Valve XV411
   		- Valve[9] : XV421 Valve XV421
   		- Valve[10]: XV431 Valve XV431
   		- Valve[11]: XV441 Valve XV441
   		- Valve[12]: XV501 Valve XV501
   		- Valve[13]: XV502 Valve XV502
   		- Valve[14]: XV901 Valve XV901
   		- Valve[15]: XV403 Valve XV403
   		- Valve[16]: XV404 Valve XV404
   		- Valve[17]: XV405 Valve XV405
   		- Valve[18]: XV406 Valve XV406
   		- Valve[19]: XV006 Valve XV006
   		- Valve[20]: XV007 Valve XV007
   		- Reset Loop : Set to 0 the Valve[21 to 99].EnableCfg
   
   -----------------------------------------------------------------------------------------------------------------------------------------------------
   	History
   		2019-AUG-13 - ACTEMIUM - B. Roch - Initial version for Candidate Release 3.00.00.00.a
   		2019-SEP-26 - ACTEMIUM - B. Roch - Modifications for Candidate Release 3.00.00.00.c
   					- Change FailState to 0 for XV441
   					- Change to valve[8] instead of Valve[0] for XV411
   		2020-SEP-30 - Merck - Q.Spindler - Modifications for Candidate Release 3.00.00.01.a
   					- Add Valves for Closed flowpath
   ============================================================*)
   
   
   (*Max valve number use as terminal value in loop
   ============================================================*)
   ValveControl.MaxValveNum := 32;
   
   (*Valve[0] : XV001 Valve XV001 (NO)
   ============================================================*)
   Valve[0].EnableCfg := 1 ;
   Valve[0].FailState := 1 ;
   Valve[0].ZSOverride := 1 ;
   Valve[0].Ports := 0 ;
   Valve[0].PriorityCfg := 0 ;
   Valve[0].ZSOpenEnable := 0 ;
   Valve[0].Alarm := 0 ;
   Valve[0].ZSCloseEnable := 0 ;
   Valve[0].ZSOpenAddress := 0 ;
   Valve[0].ZSCloseAddress := 0 ;
   Valve[0].OutputAddress := 32 ;
   
   (*Valve[1] : XV002 Valve XV002 (NO)
   ============================================================*)
   Valve[1].EnableCfg := 1 ;
   Valve[1].FailState := 1 ;
   Valve[1].ZSOverride := 1 ;
   Valve[1].Ports := 0 ;
   Valve[1].PriorityCfg := 0 ;
   Valve[1].ZSOpenEnable := 0 ;
   Valve[1].Alarm := 0 ;
   Valve[1].ZSCloseEnable := 0 ;
   Valve[1].ZSOpenAddress := 0 ;
   Valve[1].ZSCloseAddress := 0 ;
   Valve[1].OutputAddress := 33 ;
   
   (*Valve[2] : XV003 Valve XV003
   ============================================================*)
   Valve[2].EnableCfg := 1 ;
   Valve[2].FailState := 0 ;
   Valve[2].ZSOverride := 1 ;
   Valve[2].Ports := 0 ;
   Valve[2].PriorityCfg := 0 ;
   Valve[2].ZSOpenEnable := 0 ;
   Valve[2].Alarm := 0 ;
   Valve[2].ZSCloseEnable := 0 ;
   Valve[2].ZSOpenAddress := 0 ;
   Valve[2].ZSCloseAddress := 0 ;
   Valve[2].OutputAddress := 34 ;
   
   (*Valve[3] : XV004 Valve XV004
   ============================================================*)
   Valve[3].EnableCfg := 1 ;
   Valve[3].FailState := 1 ;
   Valve[3].ZSOverride := 1 ;
   Valve[3].Ports := 0 ;
   Valve[3].PriorityCfg := 0 ;
   Valve[3].ZSOpenEnable := 0 ;
   Valve[3].Alarm := 0 ;
   Valve[3].ZSCloseEnable := 0 ;
   Valve[3].ZSOpenAddress := 0 ;
   Valve[3].ZSCloseAddress := 0 ;
   Valve[3].OutputAddress := 35 ;
   
   (*Valve[4] : XV005 Valve XV005
   ============================================================*)
   Valve[4].EnableCfg := 1 ;
   Valve[4].FailState := 0 ;
   Valve[4].ZSOverride := 1 ;
   Valve[4].Ports := 0 ;
   Valve[4].PriorityCfg := 0 ;
   Valve[4].ZSOpenEnable := 0 ;
   Valve[4].Alarm := 0 ;
   Valve[4].ZSCloseEnable := 0 ;
   Valve[4].ZSOpenAddress := 0 ;
   Valve[4].ZSCloseAddress := 0 ;
   Valve[4].OutputAddress := 36 ;
   
   (*Valve[5] : XV102 Valve XV102
   ============================================================*)
   Valve[5].EnableCfg := 1 ;
   Valve[5].FailState := 0 ;
   Valve[5].ZSOverride := 1 ;
   Valve[5].Ports := 0 ;
   Valve[5].PriorityCfg := 0 ;
   Valve[5].ZSOpenEnable := 0 ;
   Valve[5].Alarm := 0 ;
   Valve[5].ZSCloseEnable := 0 ;
   Valve[5].ZSOpenAddress := 0 ;
   Valve[5].ZSCloseAddress := 0 ;
   Valve[5].OutputAddress := 38 ;
   
   (*Valve[6] : XV401 Valve XV401
   ============================================================*)
   Valve[6].EnableCfg := 1 ;
   Valve[6].FailState := 0 ;
   Valve[6].ZSOverride := 1 ;
   Valve[6].Ports := 0 ;
   Valve[6].PriorityCfg := 0 ;
   Valve[6].ZSOpenEnable := 0 ;
   Valve[6].Alarm := 0 ;
   Valve[6].ZSCloseEnable := 0 ;
   Valve[6].ZSOpenAddress := 0;
   Valve[6].ZSCloseAddress := 0 ;
   Valve[6].OutputAddress := 41 ;
   
   (*Valve[7] : XV402 Valve XV402
   ============================================================*)
   Valve[7].EnableCfg := 1 ;
   Valve[7].FailState := 0 ;
   Valve[7].ZSOverride := 1 ;
   Valve[7].Ports := 0 ;
   Valve[7].PriorityCfg := 0 ;
   Valve[7].ZSOpenEnable := 0 ;
   Valve[7].Alarm := 0 ;
   Valve[7].ZSCloseEnable := 0 ;
   Valve[7].ZSOpenAddress := 0 ;
   Valve[7].ZSCloseAddress := 0 ;
   Valve[7].OutputAddress := 42 ;
   
   (*Valve[8] : XV411 Valve XV411
   ============================================================*)
   Valve[8].EnableCfg := 1 ;
   Valve[8].FailState := 0 ;
   Valve[8].ZSOverride := 1 ;
   Valve[8].Ports := 0 ;
   Valve[8].PriorityCfg := 0 ;
   Valve[8].ZSOpenEnable := 0 ;
   Valve[8].Alarm := 0 ;
   Valve[8].ZSCloseEnable := 0 ;
   Valve[8].ZSOpenAddress := 0 ;
   Valve[8].ZSCloseAddress := 0 ;
   Valve[8].OutputAddress := 43 ;
   
   (*Valve[9] : XV421 Valve XV421
   ============================================================*)
   Valve[9].EnableCfg := 1 ;
   Valve[9].FailState := 0 ;
   Valve[9].ZSOverride := 1 ;
   Valve[9].Ports := 0 ;
   Valve[9].PriorityCfg := 0 ;
   Valve[9].ZSOpenEnable := 0 ;
   Valve[9].Alarm := 0 ;
   Valve[9].ZSCloseEnable := 0 ;
   Valve[9].ZSOpenAddress := 0 ;
   Valve[9].ZSCloseAddress := 0 ;
   Valve[9].OutputAddress := 44 ;
   
   (*Valve[10]: XV431 Valve XV431
   ============================================================*)
   Valve[10].EnableCfg := 1 ;
   Valve[10].FailState := 0 ;
   Valve[10].ZSOverride := 1 ;
   Valve[10].Ports := 0 ;
   Valve[10].PriorityCfg := 0 ;
   Valve[10].ZSOpenEnable := 0 ;
   Valve[10].Alarm := 0 ;
   Valve[10].ZSCloseEnable := 0 ;
   Valve[10].ZSOpenAddress := 0 ;
   Valve[10].ZSCloseAddress := 0 ;
   Valve[10].OutputAddress := 45 ;
   
   (*Valve[11]: XV441 Valve XV441
   ============================================================*)
   Valve[11].EnableCfg := 1 ;
   Valve[11].FailState := 0 ;
   Valve[11].ZSOverride := 1 ;
   Valve[11].Ports := 0 ;
   Valve[11].PriorityCfg := 0 ;
   Valve[11].ZSOpenEnable := 0 ;
   Valve[11].Alarm := 0 ;
   Valve[11].ZSCloseEnable := 0 ;
   Valve[11].ZSOpenAddress := 0 ;
   Valve[11].ZSCloseAddress := 0 ;
   Valve[11].OutputAddress := 46 ;
   
   (*Valve[12]: XV501 Valve XV501
   ============================================================*)
   
   IF Options.TF3S THEN
   	Valve[12].EnableCfg := 1 ;
   ELSE
   	Valve[12].EnableCfg := 0 ;
   END_IF;
   
   Valve[12].FailState := 0 ;
   Valve[12].ZSOverride := 1 ;
   Valve[12].Ports := 0 ;
   Valve[12].PriorityCfg := 0 ;
   Valve[12].ZSOpenEnable := 0 ;
   Valve[12].Alarm := 0 ;
   Valve[12].ZSCloseEnable := 0 ;
   Valve[12].ZSOpenAddress := 0 ;
   Valve[12].ZSCloseAddress := 0 ;
   Valve[12].OutputAddress := 39 ;
   
   (*Valve[13]: XV502 Valve XV502
   ============================================================*)
   
   IF Options.TF3S THEN
   	Valve[13].EnableCfg := 1 ;
   ELSE
   	Valve[13].EnableCfg := 0 ;
   END_IF;
   
   Valve[13].FailState := 0 ;
   Valve[13].ZSOverride := 1 ;
   Valve[13].Ports := 0 ;
   Valve[13].PriorityCfg := 0 ;
   Valve[13].ZSOpenEnable := 0 ;
   Valve[13].Alarm := 0 ;
   Valve[13].ZSCloseEnable := 0 ;
   Valve[13].ZSOpenAddress := 0 ;
   Valve[13].ZSCloseAddress := 0 ;
   Valve[13].OutputAddress := 40 ;
   
   (*Valve[14]: XV901 Valve XV901
   ============================================================*)
   Valve[14].EnableCfg := 1 ;
   Valve[14].FailState := 0 ;
   Valve[14].ZSOverride := 1 ;
   Valve[14].Ports := 0 ;
   Valve[14].PriorityCfg := 0 ;
   Valve[14].ZSOpenEnable := 0 ;
   Valve[14].Alarm := 0 ;
   Valve[14].ZSCloseEnable := 0 ;
   Valve[14].ZSOpenAddress := 0 ;
   Valve[14].ZSCloseAddress := 0 ;
   Valve[14].OutputAddress := 37 ;
   
   (*Valve[15]: XV403 Valve XV403
   ============================================================*)
   IF Options.ClosedFP THEN
   	Valve[15].EnableCfg := 1 ;
   ELSE
   	Valve[15].EnableCfg := 0 ;
   END_IF;
   Valve[15].FailState := 0 ;
   Valve[15].ZSOverride := 1 ;
   Valve[15].Ports := 0 ;
   Valve[15].PriorityCfg := 0 ;
   Valve[15].ZSOpenEnable := 0 ;
   Valve[15].Alarm := 0 ;
   Valve[15].ZSCloseEnable := 0 ;
   Valve[15].ZSOpenAddress := 0 ;
   Valve[15].ZSCloseAddress := 0 ;
   Valve[15].OutputAddress := 47 ;
   
   (*Valve[16]: XV404 Valve XV404
   ============================================================*)
   IF Options.ClosedFP THEN
   	Valve[16].EnableCfg := 1 ;
   ELSE
   	Valve[16].EnableCfg := 0 ;
   END_IF;
   Valve[16].FailState := 0 ;
   Valve[16].ZSOverride := 1 ;
   Valve[16].Ports := 0 ;
   Valve[16].PriorityCfg := 0 ;
   Valve[16].ZSOpenEnable := 0 ;
   Valve[16].Alarm := 0 ;
   Valve[16].ZSCloseEnable := 0 ;
   Valve[16].ZSOpenAddress := 0 ;
   Valve[16].ZSCloseAddress := 0 ;
   Valve[16].OutputAddress := 48 ;
   
   (*Valve[17]: XV405 Valve XV405
   ============================================================*)
   IF Options.ClosedFP THEN
   	Valve[17].EnableCfg := 1 ;
   ELSE
   	Valve[17].EnableCfg := 0 ;
   END_IF;
   Valve[17].FailState := 0 ;
   Valve[17].ZSOverride := 1 ;
   Valve[17].Ports := 0 ;
   Valve[17].PriorityCfg := 0 ;
   Valve[17].ZSOpenEnable := 0 ;
   Valve[17].Alarm := 0 ;
   Valve[17].ZSCloseEnable := 0 ;
   Valve[17].ZSOpenAddress := 0 ;
   Valve[17].ZSCloseAddress := 0 ;
   Valve[17].OutputAddress := 49 ;
   
   (*Valve[18]: XV406 Valve XV406
   ============================================================*)
   IF Options.ClosedFP THEN
   	Valve[18].EnableCfg := 1 ;
   ELSE
   	Valve[18].EnableCfg := 0 ;
   END_IF;
   Valve[18].FailState := 0 ;
   Valve[18].ZSOverride := 1 ;
   Valve[18].Ports := 0 ;
   Valve[18].PriorityCfg := 0 ;
   Valve[18].ZSOpenEnable := 0 ;
   Valve[18].Alarm := 0 ;
   Valve[18].ZSCloseEnable := 0 ;
   Valve[18].ZSOpenAddress := 0 ;
   Valve[18].ZSCloseAddress := 0 ;
   Valve[18].OutputAddress := 50 ;
   
   (*Valve[19]: XV006 Valve XV006
   ============================================================*)
   IF Options.ClosedFP THEN
   	Valve[19].EnableCfg := 1 ;
   ELSE
   	Valve[19].EnableCfg := 0 ;
   END_IF;
   Valve[19].FailState := 1 ;
   Valve[19].ZSOverride := 1 ;
   Valve[19].Ports := 0 ;
   Valve[19].PriorityCfg := 0 ;
   Valve[19].ZSOpenEnable := 0 ;
   Valve[19].Alarm := 0 ;
   Valve[19].ZSCloseEnable := 0 ;
   Valve[19].ZSOpenAddress := 0 ;
   Valve[19].ZSCloseAddress := 0 ;
   Valve[19].OutputAddress := 51 ;
   
   (*Valve[20]: XV007 Valve XV007
   ============================================================*)
   IF Options.ClosedFP THEN
   	Valve[20].EnableCfg := 1 ;
   ELSE
   	Valve[20].EnableCfg := 0 ;
   END_IF;
   Valve[20].FailState := 0 ;
   Valve[20].ZSOverride := 1 ;
   Valve[20].Ports := 0 ;
   Valve[20].PriorityCfg := 0 ;
   Valve[20].ZSOpenEnable := 0 ;
   Valve[20].Alarm := 0 ;
   Valve[20].ZSCloseEnable := 0 ;
   Valve[20].ZSOpenAddress := 0 ;
   Valve[20].ZSCloseAddress := 0 ;
   Valve[20].OutputAddress := 52 ;
   
   
   (*Reset Loop : Set to 0 the Valve[21 to 99].EnableCfg
   ============================================================*)
   FOR Config.IndeXValve := 21 to 99 by 1 do
   	Valve[Config.IndeXValve].EnableCfg := 0 ;
   	Valve[Config.IndeXValve].Alarm := 0 ;
   	Valve[Config.IndeXValve].Control := 0 ;
   	Valve[Config.IndeXValve].Auto := 0 ;
   	Valve[Config.IndeXValve].Manual := 0 ;
   	Valve[Config.IndeXValve].StatusWord := 0 ;
   	Valve[Config.IndeXValve].Status := 0 ;
   End_for ;
END_ROUTINE

ROUTINE Control_Loop   (* ladder *)
// Control Loop Routine
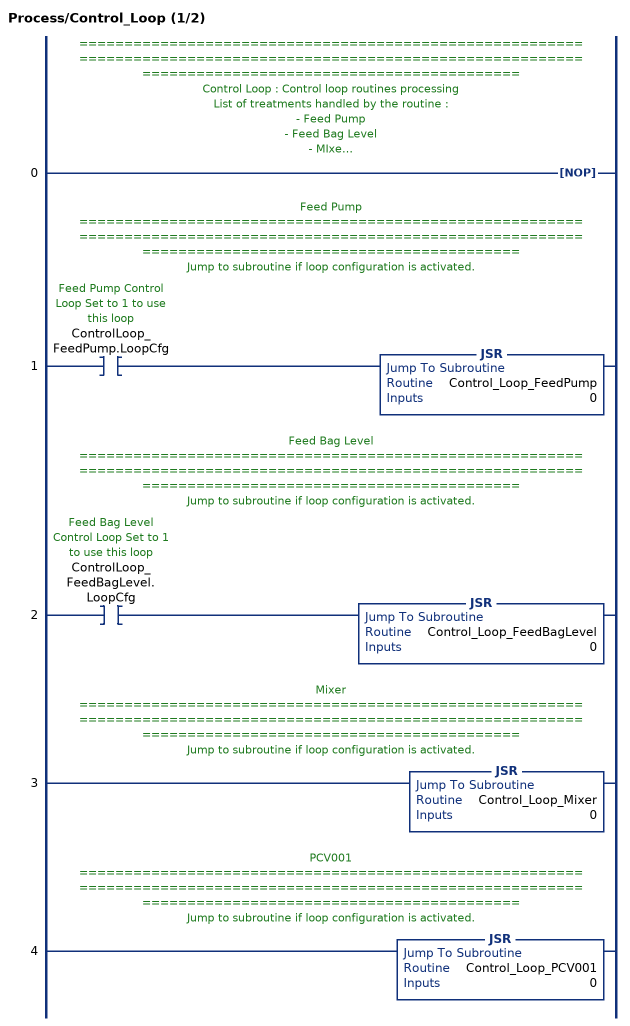
   // ==========================================================================================================================================================
   //                                                                                                                 Control Loop : Control loop routines processing
   //                                                     List of treatments handled by the routine :
   //                                                          - Feed Pump
   //                                                          - Feed Bag Level
   //                                                          - MIxer
   //                                                          - PCV001
   //                                                                                                             - PCV101                                                    -----------------------------------------------------------------------------------------------------------------------------------------------------
   //                                                     History
   //                                                         2019-AUG-13 - Actemium - B. Roch - Initial version for Candidate Release 3.00.00.00.a
   //                                                            2019-SEP-26 - Actemium - B. Roch - Initial version for Candidate Release 3.00.00.00.c
   //                                                                       - add PCV001 and PCV101 routine call
   // ==========================================================================================================================================================
   0: NOP();
   // Feed Pump
   // ==========================================================================================================================================================
   // Jump to subroutine if loop configuration is activated.
   1: XIC(ControlLoop_FeedPump.LoopCfg)JSR(Control_Loop_FeedPump,0);
   // Feed Bag Level
   // ==========================================================================================================================================================
   // Jump to subroutine if loop configuration is activated.
   2: XIC(ControlLoop_FeedBagLevel.LoopCfg)JSR(Control_Loop_FeedBagLevel,0);
   // Mixer
   // ==========================================================================================================================================================
   // Jump to subroutine if loop configuration is activated.
   3: JSR(Control_Loop_Mixer,0);
   // PCV001
   // ==========================================================================================================================================================
   // Jump to subroutine if loop configuration is activated.
   4: JSR(Control_Loop_PCV001,0);
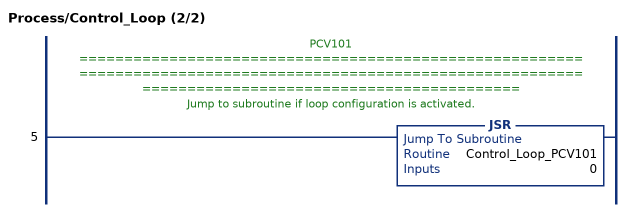
   // PCV101
   // ==========================================================================================================================================================
   // Jump to subroutine if loop configuration is activated.
   5: JSR(Control_Loop_PCV101,0);
END_ROUTINE

ROUTINE Control_Loop_FeedBagLevel   (* ladder *)
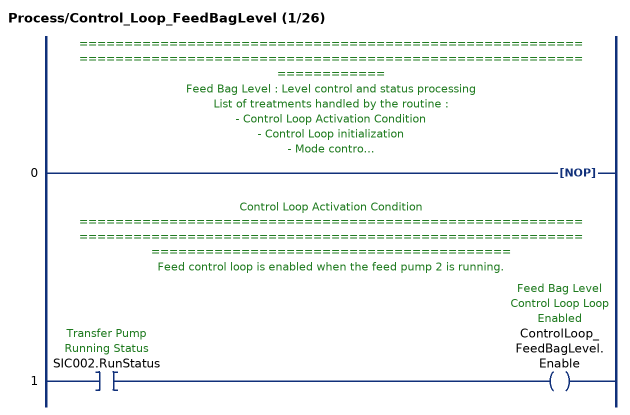
   // ============================================================================================================================
   //                                                              Feed Bag Level : Level control and status processing
   //                                                     List of treatments handled by the routine :
   //                                                          - Control Loop Activation Condition
   //                                                          - Control Loop initialization
   //                                                          - Mode control
   //                                                          - Control Loop deadband calculation
   //                                                          - Management of ramping control
   //                                                          - Control Loop Stability control
   //                                                          - Control Loop manual state control
   //                                                          - Management of PID instruction
   //                                                          - Control of the analog output
   //                                                     -----------------------------------------------------------------------------------------------------------------------------------------------------
   //                                                     History
   //    2019-AUG-13 - Actemium - B. Roch - Initial version for Candidate Release 3.00.00.00.
   //    2020-SEP-14 - Merck - Q. Spindler - Modifications for Candidate Release 3.00.00.01.a
   //                                                        - on rung 12, disable DBOK if control loop is not enabled or in manual
   // 	  2021-APR-24 - DAVIDSON- Ch. ARBOGAST - Modifications for Candidate Release 3.01.00.00.a
   // - on rung 2, line 1, replace "ControlLoop[2].Manual OR ControlLoop[2].Auto1" by
   // 			 "NOT ControlLoop[2].Auto2 AND NOT ControlLoop[2].Auto3 AND NOT ControlLoop[2].Auto4"
   // 	             - on rung 36, line 1, replace "ControlLoopFeedPump.Auto1" by "ControlLoopFeedBagLevel.Auto1"
   // ========================================================================================================================================================
   0: NOP();
   // Control Loop Activation Condition
   // ========================================================================================================================================================
   // Feed control loop is enabled when the feed pump 2 is running.
   1: XIC(SIC002.RunStatus)OTE(ControlLoop_FeedBagLevel.Enable);
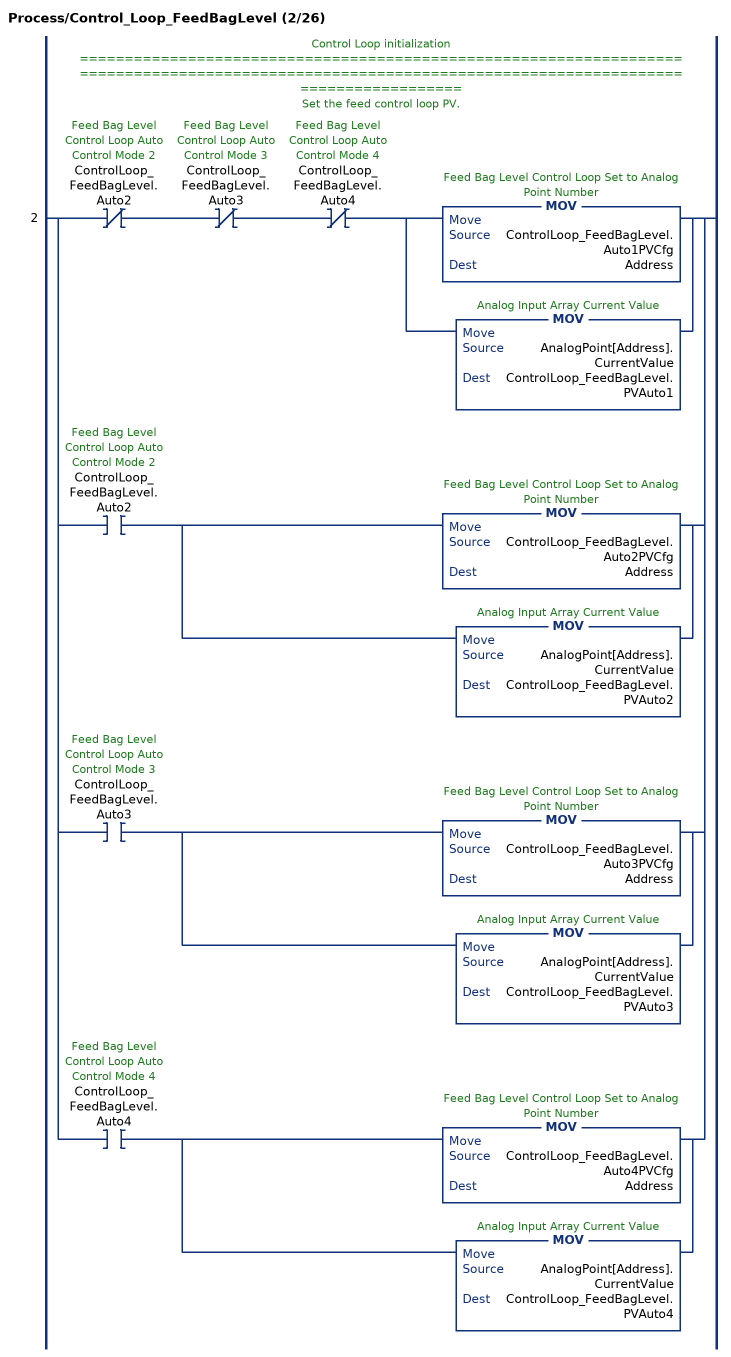
   // Control Loop initialization
   // ========================================================================================================================================================
   // Set the feed control loop PV.
   2: [[XIO(ControlLoop_FeedBagLevel.Auto2) XIO(ControlLoop_FeedBagLevel.Auto3) XIO(ControlLoop_FeedBagLevel.Auto4) [MOV(ControlLoop_FeedBagLevel.Auto1PVCfg,Address) ,MOV(AnalogPoint[Address].CurrentValue,ControlLoop_FeedBagLevel.PVAuto1) ] ,XIC(ControlLoop_FeedBagLevel.Auto2) [MOV(ControlLoop_FeedBagLevel.Auto2PVCfg,Address) ,MOV(AnalogPoint[Address].CurrentValue,ControlLoop_FeedBagLevel.PVAuto2) ] ] ,XIC(ControlLoop_FeedBagLevel.Auto3) [MOV(ControlLoop_FeedBagLevel.Auto3PVCfg,Address) ,MOV(AnalogPoint[Address].CurrentValue,ControlLoop_FeedBagLevel.PVAuto3) ] ,XIC(ControlLoop_FeedBagLevel.Auto4) [MOV(ControlLoop_FeedBagLevel.Auto4PVCfg,Address) ,MOV(AnalogPoint[Address].CurrentValue,ControlLoop_FeedBagLevel.PVAuto4) ] ];
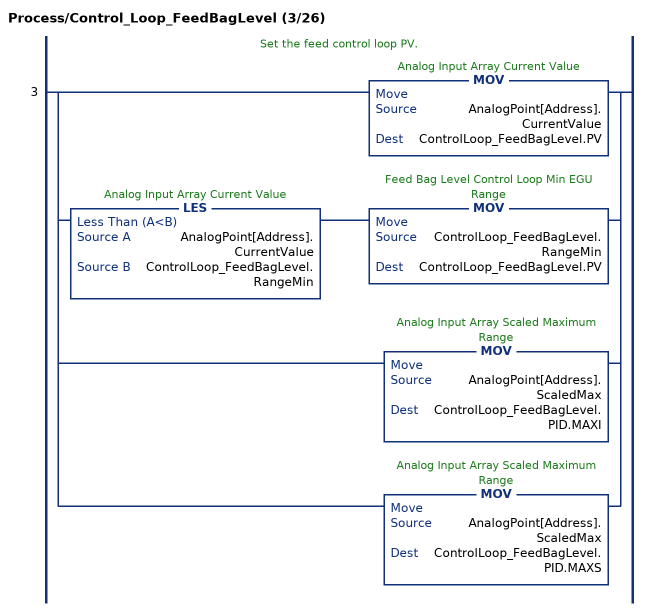
   // Set the feed control loop PV.
   3: [MOV(AnalogPoint[Address].CurrentValue,ControlLoop_FeedBagLevel.PV) ,LES(AnalogPoint[Address].CurrentValue,ControlLoop_FeedBagLevel.RangeMin) MOV(ControlLoop_FeedBagLevel.RangeMin,ControlLoop_FeedBagLevel.PV) ,MOV(AnalogPoint[Address].ScaledMax,ControlLoop_FeedBagLevel.PID.MAXI) ,MOV(AnalogPoint[Address].ScaledMax,ControlLoop_FeedBagLevel.PID.MAXS) ];
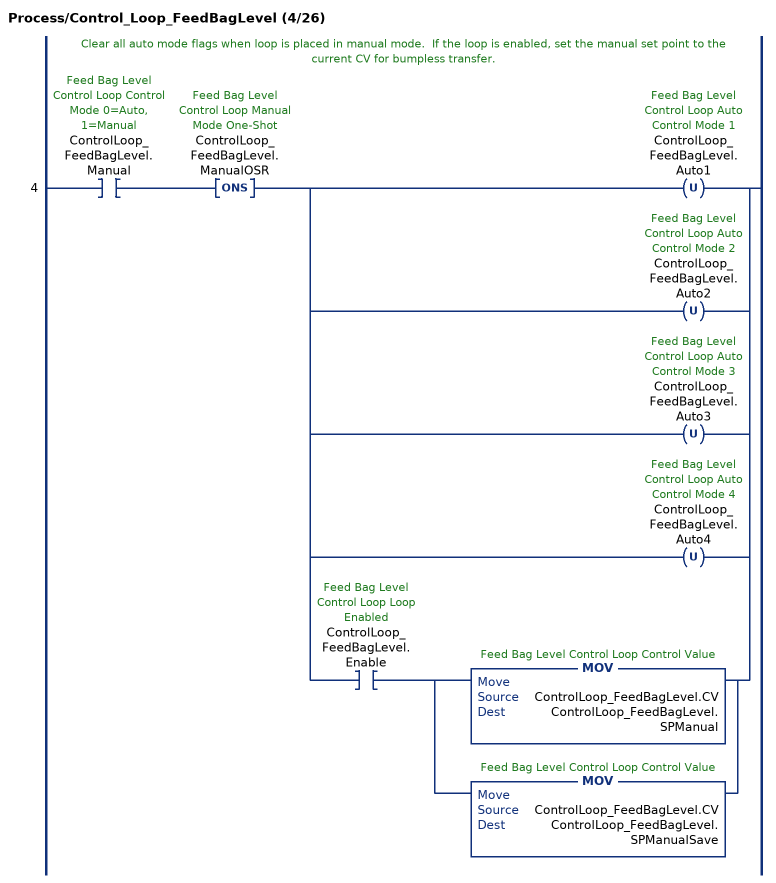
   // Clear all auto mode flags when loop is placed in manual mode.  If the loop is enabled, set the manual set point to the current CV for bumpless transfer.
   4: XIC(ControlLoop_FeedBagLevel.Manual)ONS(ControlLoop_FeedBagLevel.ManualOSR)[OTU(ControlLoop_FeedBagLevel.Auto1) ,OTU(ControlLoop_FeedBagLevel.Auto2) ,OTU(ControlLoop_FeedBagLevel.Auto3) ,OTU(ControlLoop_FeedBagLevel.Auto4) ,XIC(ControlLoop_FeedBagLevel.Enable) [MOV(ControlLoop_FeedBagLevel.CV,ControlLoop_FeedBagLevel.SPManual) ,MOV(ControlLoop_FeedBagLevel.CV,ControlLoop_FeedBagLevel.SPManualSave) ] ];
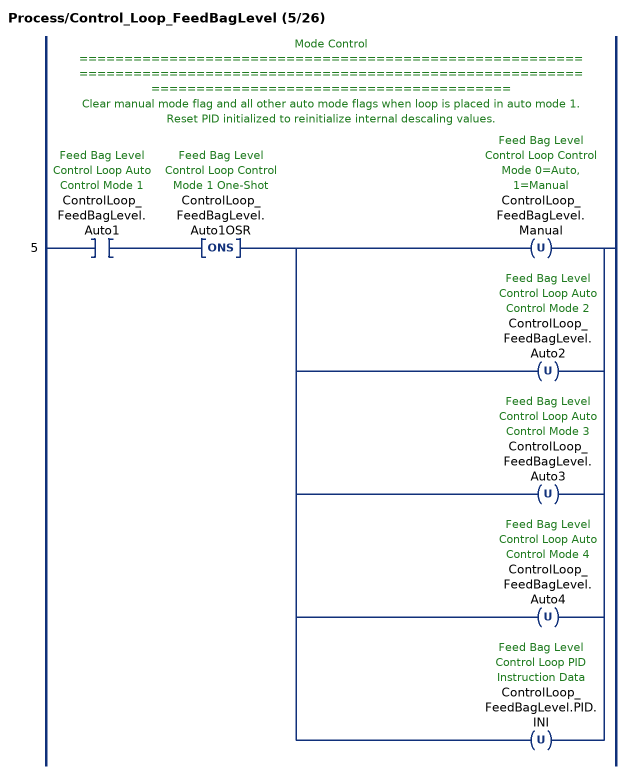
   // Mode Control
   // ========================================================================================================================================================
   // Clear manual mode flag and all other auto mode flags when loop is placed in auto mode 1. Reset PID initialized to reinitialize internal descaling values.
   5: XIC(ControlLoop_FeedBagLevel.Auto1)ONS(ControlLoop_FeedBagLevel.Auto1OSR)[OTU(ControlLoop_FeedBagLevel.Manual) ,OTU(ControlLoop_FeedBagLevel.Auto2) ,OTU(ControlLoop_FeedBagLevel.Auto3) ,OTU(ControlLoop_FeedBagLevel.Auto4) ,OTU(ControlLoop_FeedBagLevel.PID.INI) ];
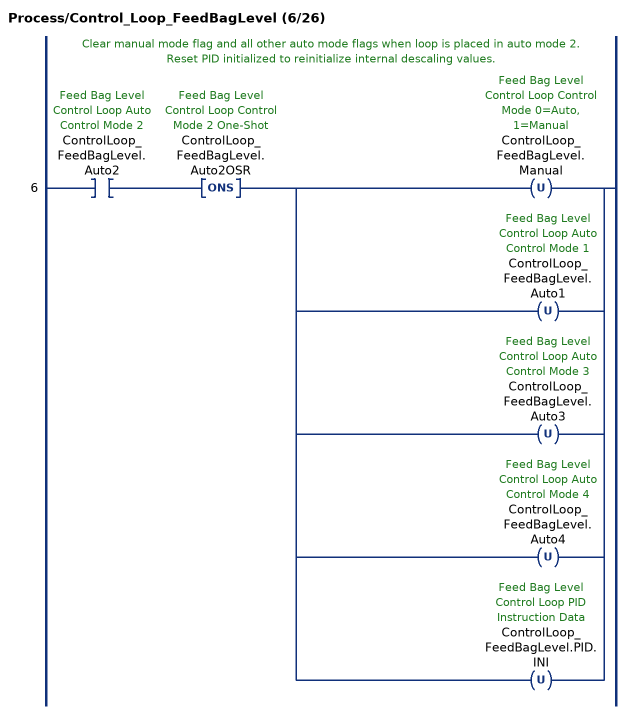
   // Clear manual mode flag and all other auto mode flags when loop is placed in auto mode 2. Reset PID initialized to reinitialize internal descaling values.
   6: XIC(ControlLoop_FeedBagLevel.Auto2)ONS(ControlLoop_FeedBagLevel.Auto2OSR)[OTU(ControlLoop_FeedBagLevel.Manual) ,OTU(ControlLoop_FeedBagLevel.Auto1) ,OTU(ControlLoop_FeedBagLevel.Auto3) ,OTU(ControlLoop_FeedBagLevel.Auto4) ,OTU(ControlLoop_FeedBagLevel.PID.INI) ];
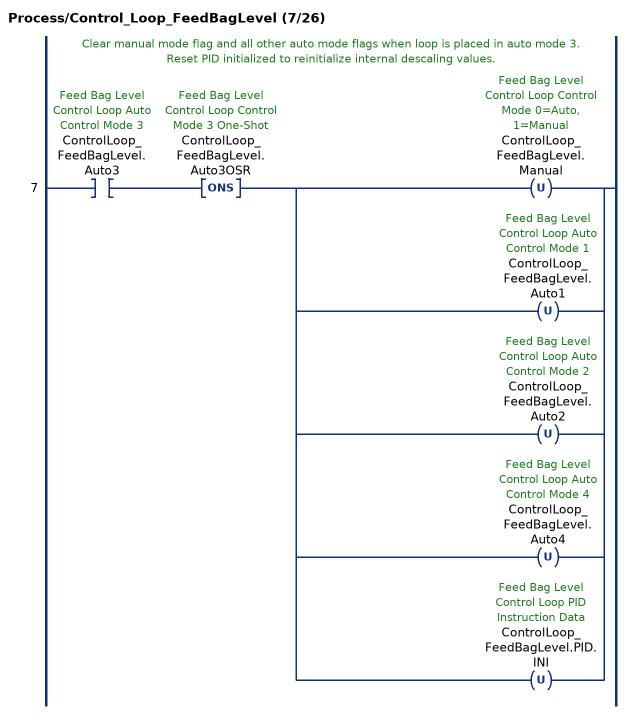
   // Clear manual mode flag and all other auto mode flags when loop is placed in auto mode 3. Reset PID initialized to reinitialize internal descaling values.
   7: XIC(ControlLoop_FeedBagLevel.Auto3)ONS(ControlLoop_FeedBagLevel.Auto3OSR)[OTU(ControlLoop_FeedBagLevel.Manual) ,OTU(ControlLoop_FeedBagLevel.Auto1) ,OTU(ControlLoop_FeedBagLevel.Auto2) ,OTU(ControlLoop_FeedBagLevel.Auto4) ,OTU(ControlLoop_FeedBagLevel.PID.INI) ];
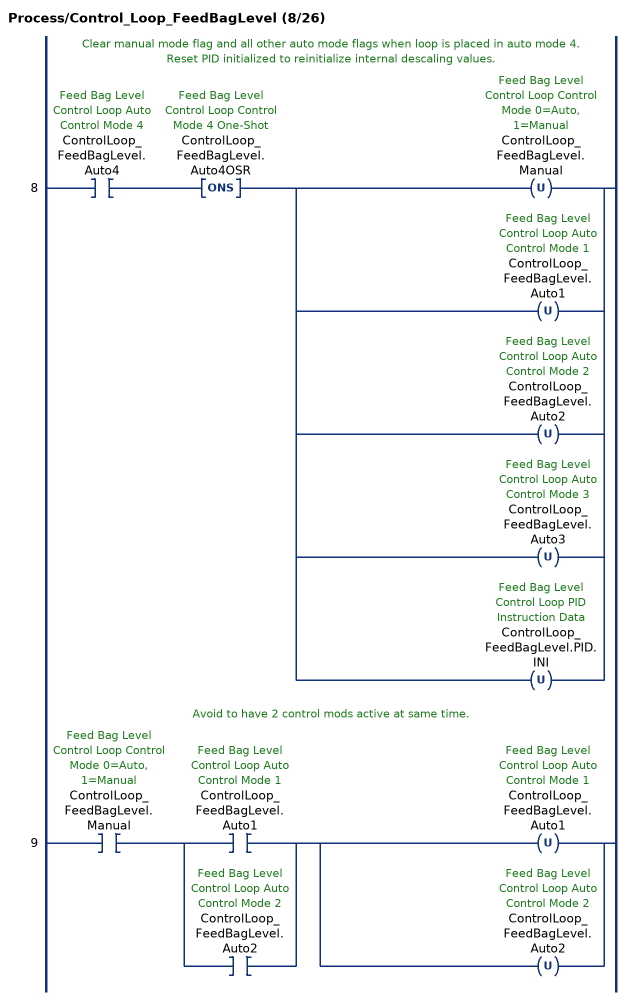
   // Clear manual mode flag and all other auto mode flags when loop is placed in auto mode 4. Reset PID initialized to reinitialize internal descaling values.
   8: XIC(ControlLoop_FeedBagLevel.Auto4)ONS(ControlLoop_FeedBagLevel.Auto4OSR)[OTU(ControlLoop_FeedBagLevel.Manual) ,OTU(ControlLoop_FeedBagLevel.Auto1) ,OTU(ControlLoop_FeedBagLevel.Auto2) ,OTU(ControlLoop_FeedBagLevel.Auto3) ,OTU(ControlLoop_FeedBagLevel.PID.INI) ];
   // Avoid to have 2 control mods active at same time.
   9: XIC(ControlLoop_FeedBagLevel.Manual)[XIC(ControlLoop_FeedBagLevel.Auto1) ,XIC(ControlLoop_FeedBagLevel.Auto2) ][OTU(ControlLoop_FeedBagLevel.Auto1) ,OTU(ControlLoop_FeedBagLevel.Auto2) ];
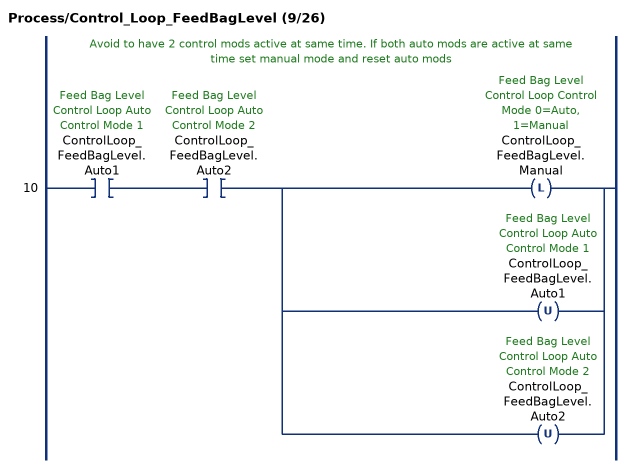
   // Avoid to have 2 control mods active at same time. If both auto mods are active at same time set manual mode and reset auto mods
   10: XIC(ControlLoop_FeedBagLevel.Auto1)XIC(ControlLoop_FeedBagLevel.Auto2)[OTL(ControlLoop_FeedBagLevel.Manual) ,OTU(ControlLoop_FeedBagLevel.Auto1) ,OTU(ControlLoop_FeedBagLevel.Auto2) ];
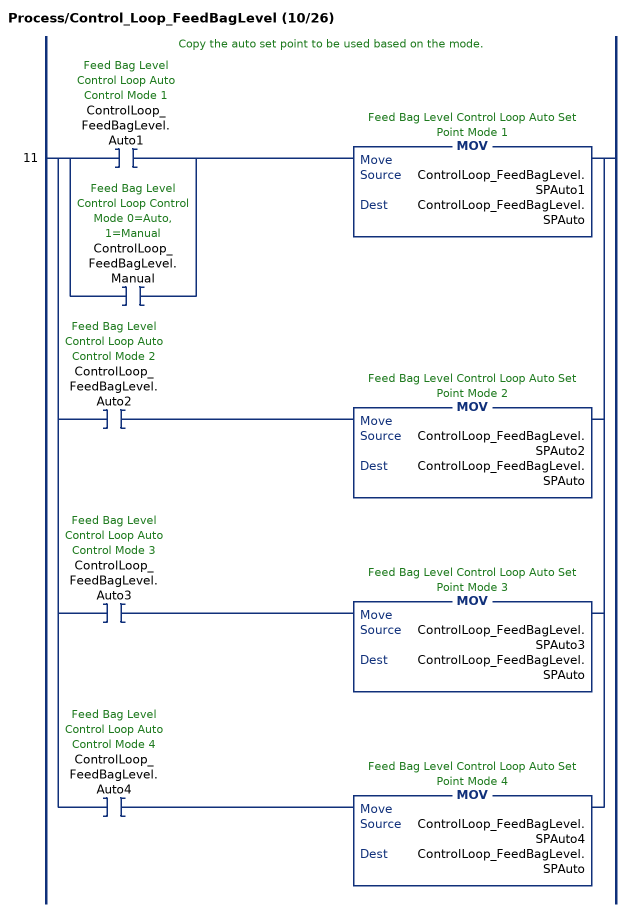
   // Copy the auto set point to be used based on the mode.
   11: [[XIC(ControlLoop_FeedBagLevel.Auto1) ,XIC(ControlLoop_FeedBagLevel.Manual) ] MOV(ControlLoop_FeedBagLevel.SPAuto1,ControlLoop_FeedBagLevel.SPAuto) ,XIC(ControlLoop_FeedBagLevel.Auto2) MOV(ControlLoop_FeedBagLevel.SPAuto2,ControlLoop_FeedBagLevel.SPAuto) ,XIC(ControlLoop_FeedBagLevel.Auto3) MOV(ControlLoop_FeedBagLevel.SPAuto3,ControlLoop_FeedBagLevel.SPAuto) ,XIC(ControlLoop_FeedBagLevel.Auto4) MOV(ControlLoop_FeedBagLevel.SPAuto4,ControlLoop_FeedBagLevel.SPAuto) ];
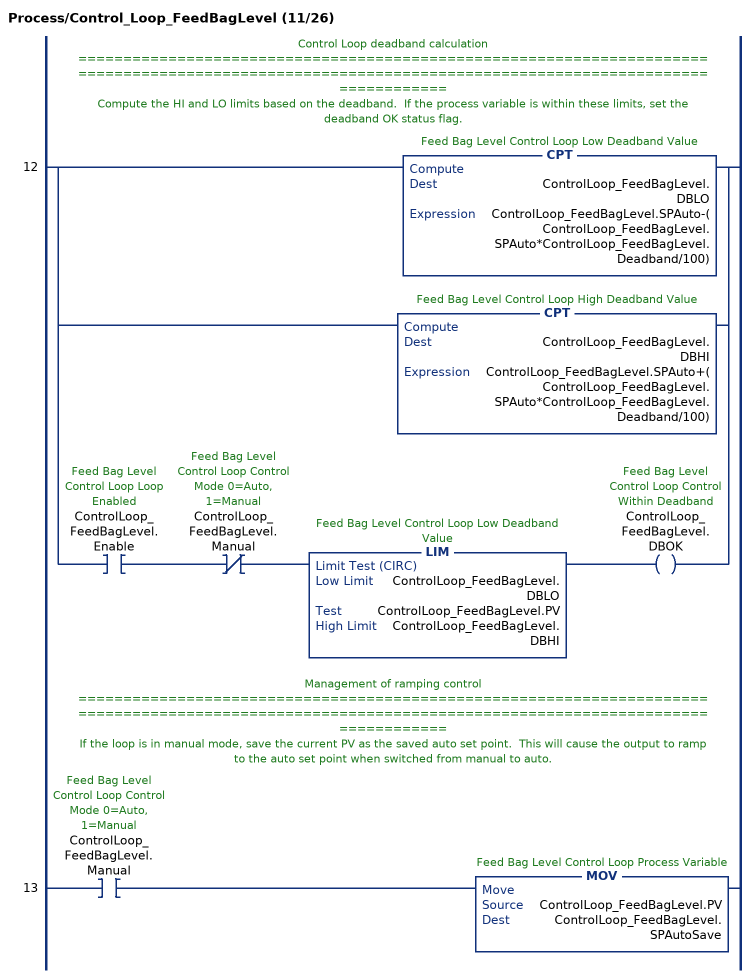
   // Control Loop deadband calculation
   // ========================================================================================================================================================
   // Compute the HI and LO limits based on the deadband.  If the process variable is within these limits, set the deadband OK status flag.
   12: [CPT(ControlLoop_FeedBagLevel.DBLO,ControlLoop_FeedBagLevel.SPAuto-(ControlLoop_FeedBagLevel.SPAuto*ControlLoop_FeedBagLevel.Deadband/100)) ,CPT(ControlLoop_FeedBagLevel.DBHI,ControlLoop_FeedBagLevel.SPAuto+(ControlLoop_FeedBagLevel.SPAuto*ControlLoop_FeedBagLevel.Deadband/100)) ,XIC(ControlLoop_FeedBagLevel.Enable) XIO(ControlLoop_FeedBagLevel.Manual) LIM(ControlLoop_FeedBagLevel.DBLO,ControlLoop_FeedBagLevel.PV,ControlLoop_FeedBagLevel.DBHI) OTE(ControlLoop_FeedBagLevel.DBOK) ];
   // Management of ramping control
   // ========================================================================================================================================================
   // If the loop is in manual mode, save the current PV as the saved auto set point.  This will cause the output to ramp to the auto set point when switched from manual to auto.
   13: XIC(ControlLoop_FeedBagLevel.Manual)MOV(ControlLoop_FeedBagLevel.PV,ControlLoop_FeedBagLevel.SPAutoSave);
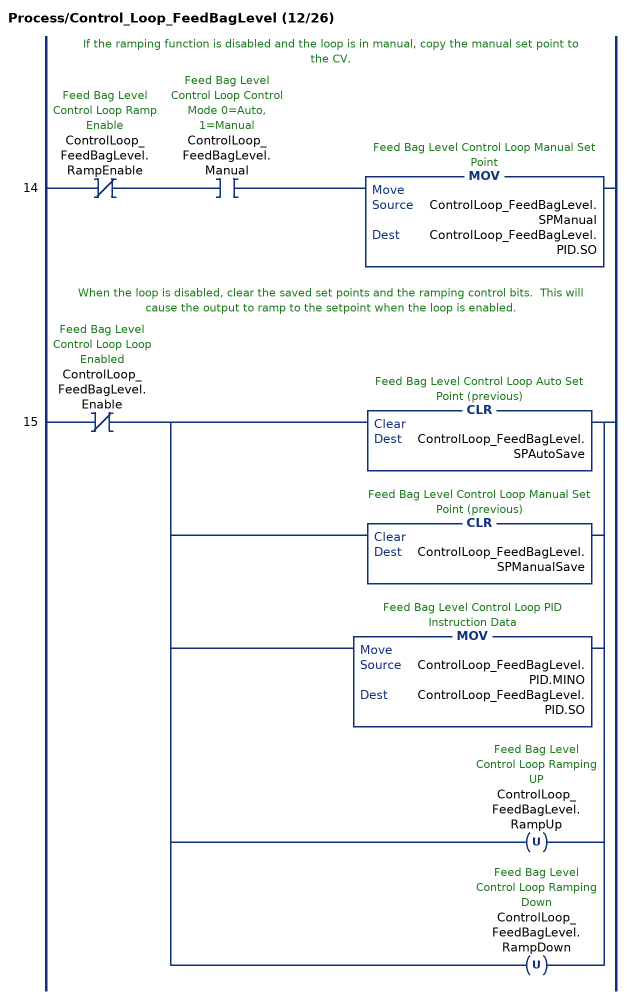
   // If the ramping function is disabled and the loop is in manual, copy the manual set point to the CV.
   14: XIO(ControlLoop_FeedBagLevel.RampEnable)XIC(ControlLoop_FeedBagLevel.Manual)MOV(ControlLoop_FeedBagLevel.SPManual,ControlLoop_FeedBagLevel.PID.SO);
   // When the loop is disabled, clear the saved set points and the ramping control bits.  This will cause the output to ramp to the setpoint when the loop is enabled.
   15: XIO(ControlLoop_FeedBagLevel.Enable)[CLR(ControlLoop_FeedBagLevel.SPAutoSave) ,CLR(ControlLoop_FeedBagLevel.SPManualSave) ,MOV(ControlLoop_FeedBagLevel.PID.MINO,ControlLoop_FeedBagLevel.PID.SO) ,OTU(ControlLoop_FeedBagLevel.RampUp) ,OTU(ControlLoop_FeedBagLevel.RampDown) ];
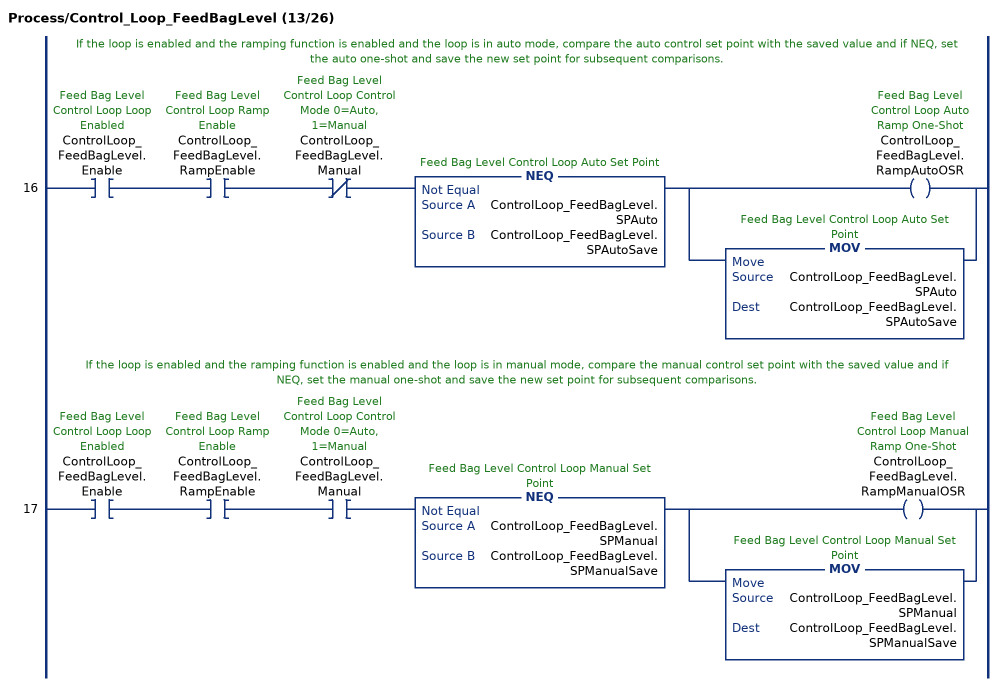
   // If the loop is enabled and the ramping function is enabled and the loop is in auto mode, compare the auto control set point with the saved value and if NEQ, set the auto one-shot and save the new set point for subsequent comparisons.
   16: XIC(ControlLoop_FeedBagLevel.Enable)XIC(ControlLoop_FeedBagLevel.RampEnable)XIO(ControlLoop_FeedBagLevel.Manual)NEQ(ControlLoop_FeedBagLevel.SPAuto,ControlLoop_FeedBagLevel.SPAutoSave)[OTE(ControlLoop_FeedBagLevel.RampAutoOSR) ,MOV(ControlLoop_FeedBagLevel.SPAuto,ControlLoop_FeedBagLevel.SPAutoSave) ];
   // If the loop is enabled and the ramping function is enabled and the loop is in manual mode, compare the manual control set point with the saved value and if NEQ, set the manual one-shot and save the new set point for subsequent comparisons.
   17: XIC(ControlLoop_FeedBagLevel.Enable)XIC(ControlLoop_FeedBagLevel.RampEnable)XIC(ControlLoop_FeedBagLevel.Manual)NEQ(ControlLoop_FeedBagLevel.SPManual,ControlLoop_FeedBagLevel.SPManualSave)[OTE(ControlLoop_FeedBagLevel.RampManualOSR) ,MOV(ControlLoop_FeedBagLevel.SPManual,ControlLoop_FeedBagLevel.SPManualSave) ];
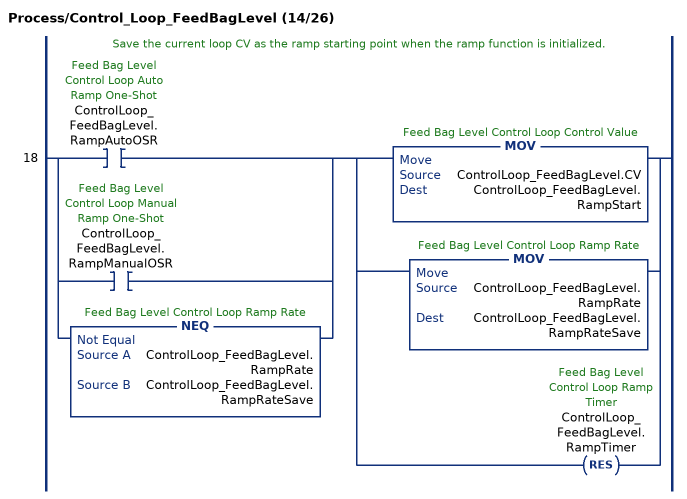
   // Save the current loop CV as the ramp starting point when the ramp function is initialized.
   18: [XIC(ControlLoop_FeedBagLevel.RampAutoOSR) ,XIC(ControlLoop_FeedBagLevel.RampManualOSR) ,NEQ(ControlLoop_FeedBagLevel.RampRate,ControlLoop_FeedBagLevel.RampRateSave) ][MOV(ControlLoop_FeedBagLevel.CV,ControlLoop_FeedBagLevel.RampStart) ,MOV(ControlLoop_FeedBagLevel.RampRate,ControlLoop_FeedBagLevel.RampRateSave) ,RES(ControlLoop_FeedBagLevel.RampTimer) ];
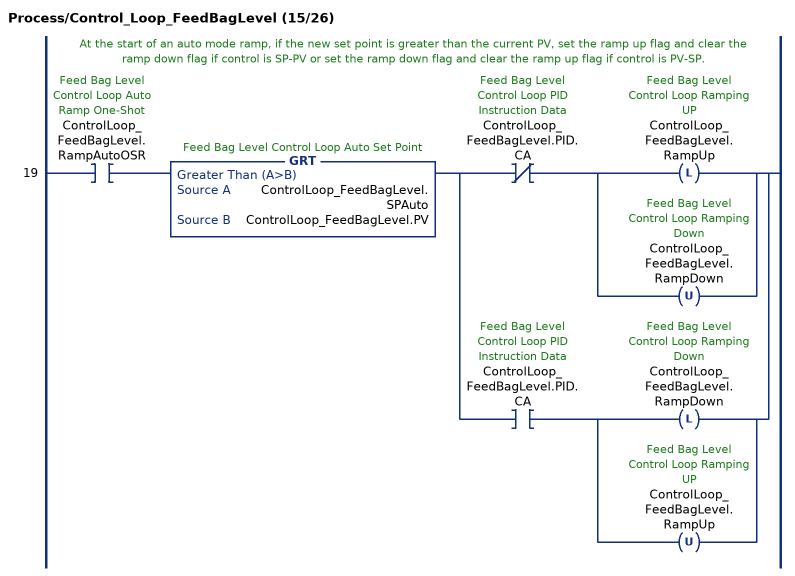
   // At the start of an auto mode ramp, if the new set point is greater than the current PV, set the ramp up flag and clear the ramp down flag if control is SP-PV or set the ramp down flag and clear the ramp up flag if control is PV-SP.
   19: XIC(ControlLoop_FeedBagLevel.RampAutoOSR)GRT(ControlLoop_FeedBagLevel.SPAuto,ControlLoop_FeedBagLevel.PV)[XIO(ControlLoop_FeedBagLevel.PID.CA) [OTL(ControlLoop_FeedBagLevel.RampUp) ,OTU(ControlLoop_FeedBagLevel.RampDown) ] ,XIC(ControlLoop_FeedBagLevel.PID.CA) [OTL(ControlLoop_FeedBagLevel.RampDown) ,OTU(ControlLoop_FeedBagLevel.RampUp) ] ];
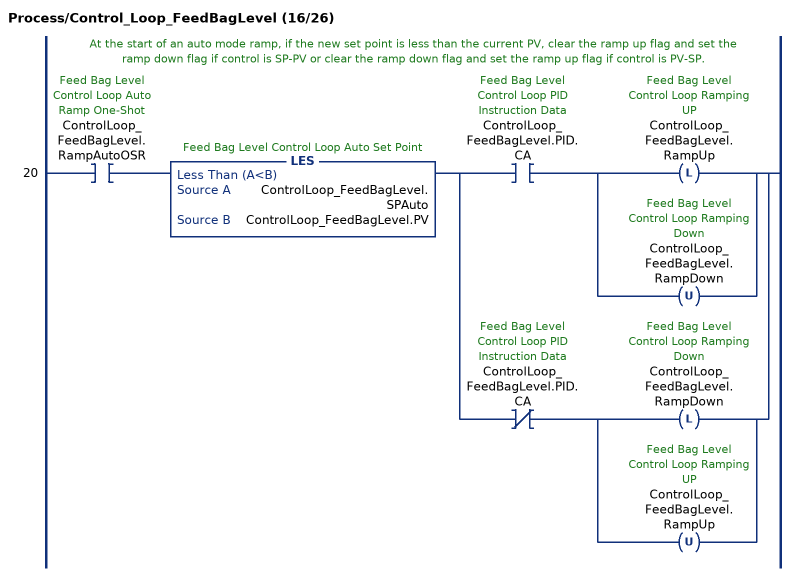
   // At the start of an auto mode ramp, if the new set point is less than the current PV, clear the ramp up flag and set the ramp down flag if control is SP-PV or clear the ramp down flag and set the ramp up flag if control is PV-SP.
   20: XIC(ControlLoop_FeedBagLevel.RampAutoOSR)LES(ControlLoop_FeedBagLevel.SPAuto,ControlLoop_FeedBagLevel.PV)[XIC(ControlLoop_FeedBagLevel.PID.CA) [OTL(ControlLoop_FeedBagLevel.RampUp) ,OTU(ControlLoop_FeedBagLevel.RampDown) ] ,XIO(ControlLoop_FeedBagLevel.PID.CA) [OTL(ControlLoop_FeedBagLevel.RampDown) ,OTU(ControlLoop_FeedBagLevel.RampUp) ] ];
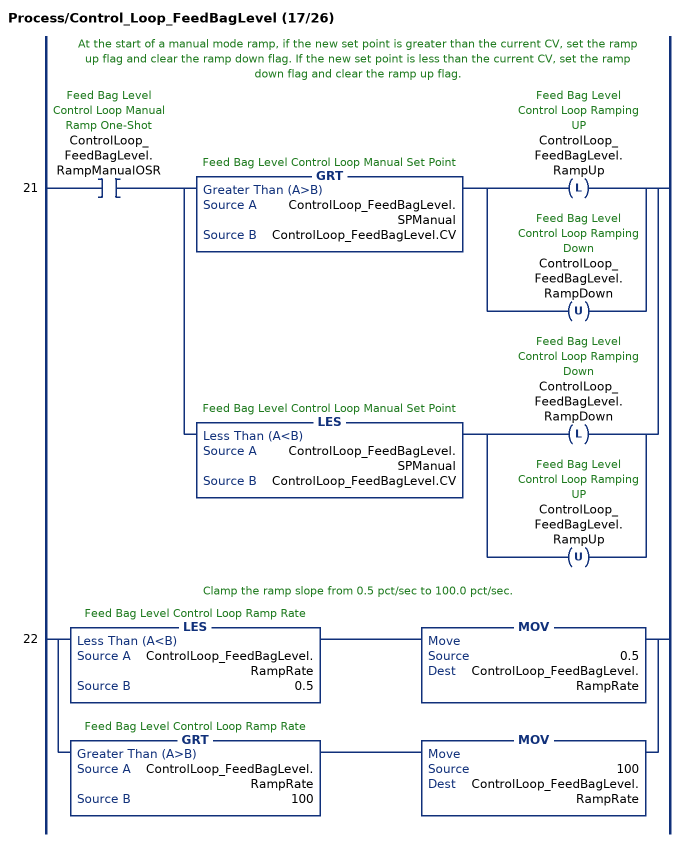
   // At the start of a manual mode ramp, if the new set point is greater than the current CV, set the ramp up flag and clear the ramp down flag. If the new set point is less than the current CV, set the ramp down flag and clear the ramp up flag.
   21: XIC(ControlLoop_FeedBagLevel.RampManualOSR)[GRT(ControlLoop_FeedBagLevel.SPManual,ControlLoop_FeedBagLevel.CV) [OTL(ControlLoop_FeedBagLevel.RampUp) ,OTU(ControlLoop_FeedBagLevel.RampDown) ] ,LES(ControlLoop_FeedBagLevel.SPManual,ControlLoop_FeedBagLevel.CV) [OTL(ControlLoop_FeedBagLevel.RampDown) ,OTU(ControlLoop_FeedBagLevel.RampUp) ] ];
   // Clamp the ramp slope from 0.5 pct/sec to 100.0 pct/sec.
   22: [LES(ControlLoop_FeedBagLevel.RampRate,0.5) MOV(0.5,ControlLoop_FeedBagLevel.RampRate) ,GRT(ControlLoop_FeedBagLevel.RampRate,100) MOV(100,ControlLoop_FeedBagLevel.RampRate) ];
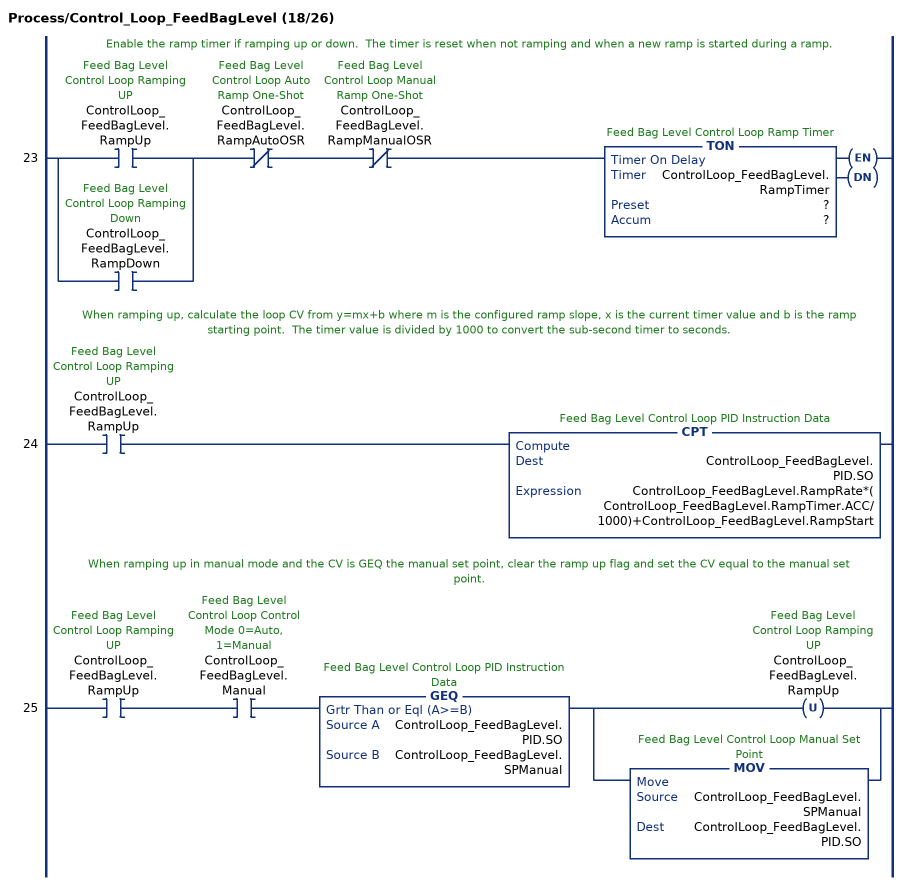
   // Enable the ramp timer if ramping up or down.  The timer is reset when not ramping and when a new ramp is started during a ramp.
   23: [XIC(ControlLoop_FeedBagLevel.RampUp) ,XIC(ControlLoop_FeedBagLevel.RampDown) ]XIO(ControlLoop_FeedBagLevel.RampAutoOSR)XIO(ControlLoop_FeedBagLevel.RampManualOSR)TON(ControlLoop_FeedBagLevel.RampTimer,?,?);
   // When ramping up, calculate the loop CV from y=mx+b where m is the configured ramp slope, x is the current timer value and b is the ramp starting point.  The timer value is divided by 1000 to convert the sub-second timer to seconds.
   24: XIC(ControlLoop_FeedBagLevel.RampUp)CPT(ControlLoop_FeedBagLevel.PID.SO,ControlLoop_FeedBagLevel.RampRate*(ControlLoop_FeedBagLevel.RampTimer.ACC/1000)+ControlLoop_FeedBagLevel.RampStart);
   // When ramping up in manual mode and the CV is GEQ the manual set point, clear the ramp up flag and set the CV equal to the manual set point.
   25: XIC(ControlLoop_FeedBagLevel.RampUp)XIC(ControlLoop_FeedBagLevel.Manual)GEQ(ControlLoop_FeedBagLevel.PID.SO,ControlLoop_FeedBagLevel.SPManual)[OTU(ControlLoop_FeedBagLevel.RampUp) ,MOV(ControlLoop_FeedBagLevel.SPManual,ControlLoop_FeedBagLevel.PID.SO) ];
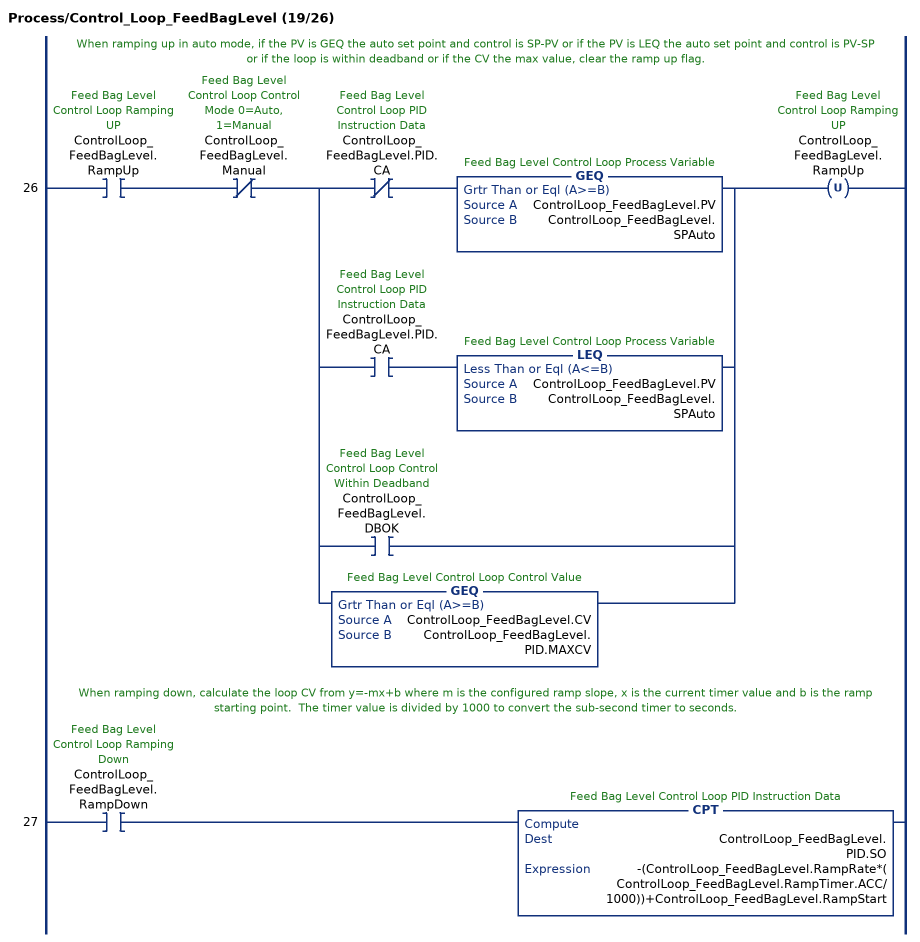
   // When ramping up in auto mode, if the PV is GEQ the auto set point and control is SP-PV or if the PV is LEQ the auto set point and control is PV-SP or if the loop is within deadband or if the CV the max value, clear the ramp up flag.
   26: XIC(ControlLoop_FeedBagLevel.RampUp)XIO(ControlLoop_FeedBagLevel.Manual)[XIO(ControlLoop_FeedBagLevel.PID.CA) GEQ(ControlLoop_FeedBagLevel.PV,ControlLoop_FeedBagLevel.SPAuto) ,XIC(ControlLoop_FeedBagLevel.PID.CA) LEQ(ControlLoop_FeedBagLevel.PV,ControlLoop_FeedBagLevel.SPAuto) ,XIC(ControlLoop_FeedBagLevel.DBOK) ,GEQ(ControlLoop_FeedBagLevel.CV,ControlLoop_FeedBagLevel.PID.MAXCV) ]OTU(ControlLoop_FeedBagLevel.RampUp);
   // When ramping down, calculate the loop CV from y=-mx+b where m is the configured ramp slope, x is the current timer value and b is the ramp starting point.  The timer value is divided by 1000 to convert the sub-second timer to seconds.
   27: XIC(ControlLoop_FeedBagLevel.RampDown)CPT(ControlLoop_FeedBagLevel.PID.SO,-(ControlLoop_FeedBagLevel.RampRate*(ControlLoop_FeedBagLevel.RampTimer.ACC/1000))+ControlLoop_FeedBagLevel.RampStart);
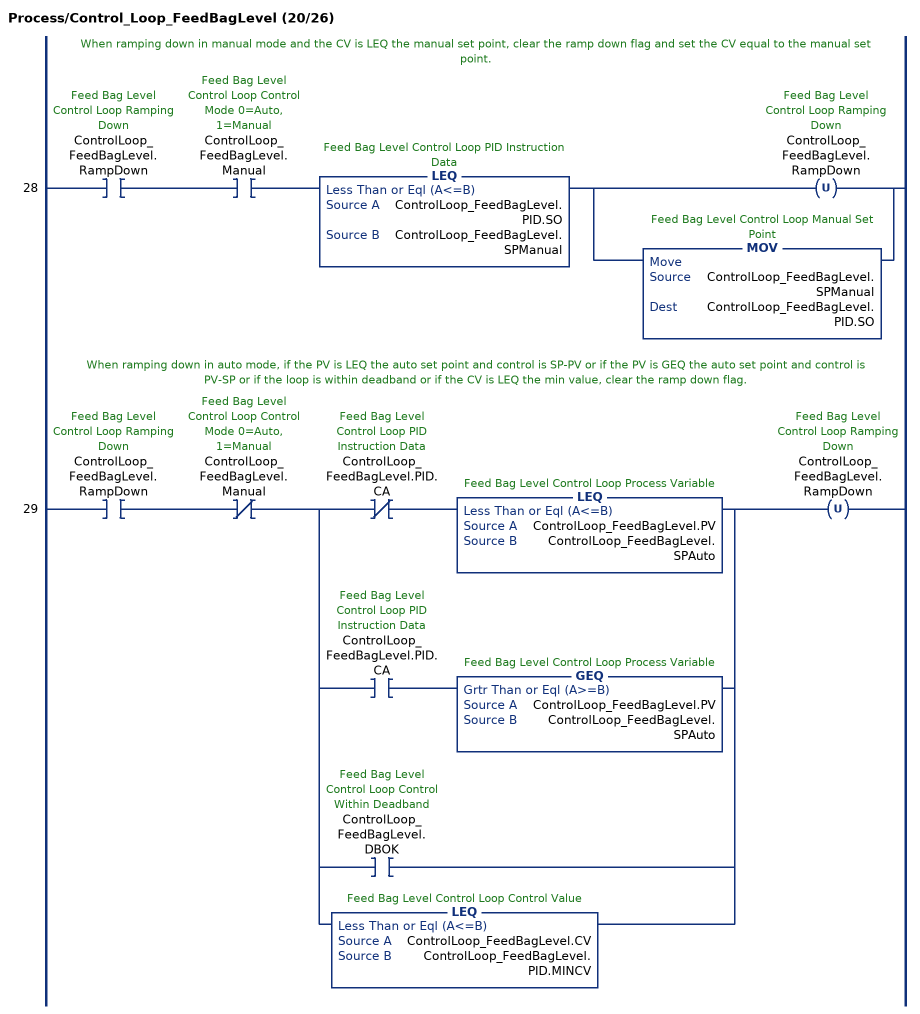
   // When ramping down in manual mode and the CV is LEQ the manual set point, clear the ramp down flag and set the CV equal to the manual set point.
   28: XIC(ControlLoop_FeedBagLevel.RampDown)XIC(ControlLoop_FeedBagLevel.Manual)LEQ(ControlLoop_FeedBagLevel.PID.SO,ControlLoop_FeedBagLevel.SPManual)[OTU(ControlLoop_FeedBagLevel.RampDown) ,MOV(ControlLoop_FeedBagLevel.SPManual,ControlLoop_FeedBagLevel.PID.SO) ];
   // When ramping down in auto mode, if the PV is LEQ the auto set point and control is SP-PV or if the PV is GEQ the auto set point and control is PV-SP or if the loop is within deadband or if the CV is LEQ the min value, clear the ramp down flag.
   29: XIC(ControlLoop_FeedBagLevel.RampDown)XIO(ControlLoop_FeedBagLevel.Manual)[XIO(ControlLoop_FeedBagLevel.PID.CA) LEQ(ControlLoop_FeedBagLevel.PV,ControlLoop_FeedBagLevel.SPAuto) ,XIC(ControlLoop_FeedBagLevel.PID.CA) GEQ(ControlLoop_FeedBagLevel.PV,ControlLoop_FeedBagLevel.SPAuto) ,XIC(ControlLoop_FeedBagLevel.DBOK) ,LEQ(ControlLoop_FeedBagLevel.CV,ControlLoop_FeedBagLevel.PID.MINCV) ]OTU(ControlLoop_FeedBagLevel.RampDown);
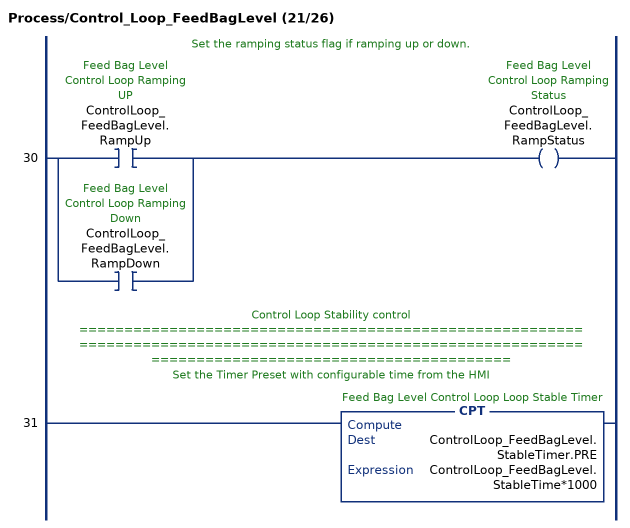
   // Set the ramping status flag if ramping up or down.
   30: [XIC(ControlLoop_FeedBagLevel.RampUp) ,XIC(ControlLoop_FeedBagLevel.RampDown) ]OTE(ControlLoop_FeedBagLevel.RampStatus);
   // Control Loop Stability control
   // ========================================================================================================================================================
   // Set the Timer Preset with configurable time from the HMI
   31: CPT(ControlLoop_FeedBagLevel.StableTimer.PRE,ControlLoop_FeedBagLevel.StableTime*1000);
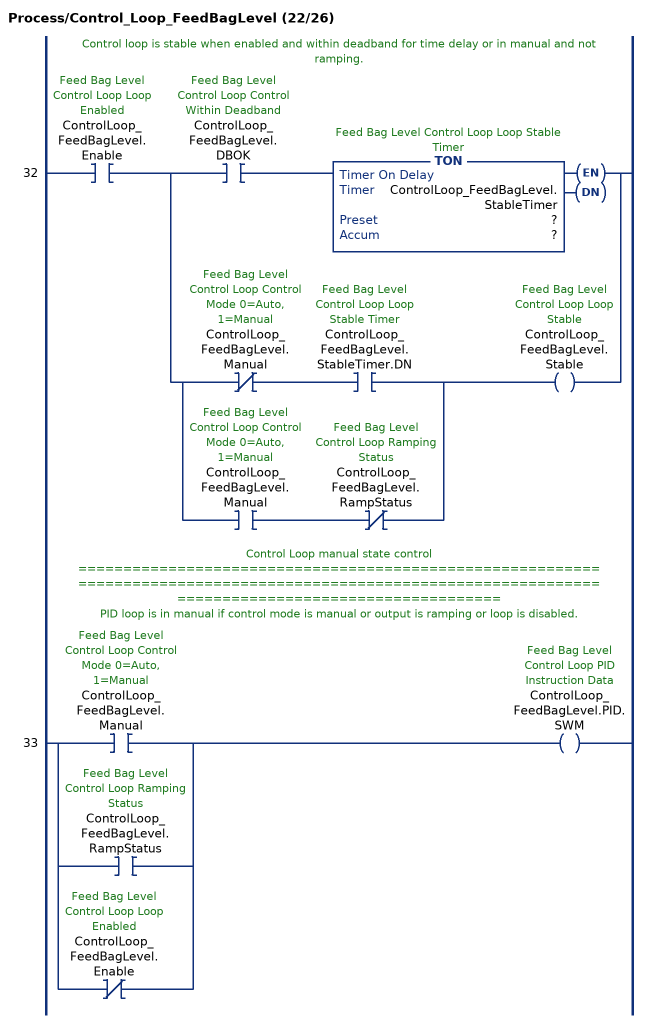
   // Control loop is stable when enabled and within deadband for time delay or in manual and not ramping.
   32: XIC(ControlLoop_FeedBagLevel.Enable)[XIC(ControlLoop_FeedBagLevel.DBOK) TON(ControlLoop_FeedBagLevel.StableTimer,?,?) ,[XIO(ControlLoop_FeedBagLevel.Manual) XIC(ControlLoop_FeedBagLevel.StableTimer.DN) ,XIC(ControlLoop_FeedBagLevel.Manual) XIO(ControlLoop_FeedBagLevel.RampStatus) ] OTE(ControlLoop_FeedBagLevel.Stable) ];
   // Control Loop manual state control
   // ========================================================================================================================================================
   // PID loop is in manual if control mode is manual or output is ramping or loop is disabled.
   33: [XIC(ControlLoop_FeedBagLevel.Manual) ,XIC(ControlLoop_FeedBagLevel.RampStatus) ,XIO(ControlLoop_FeedBagLevel.Enable) ]OTE(ControlLoop_FeedBagLevel.PID.SWM);
